(* CODESYS project process.library
   DefaultNamespace: KOSTAL.TC3.Core.process
   Description: Core Functionalities
   Author: Frank Dümpelmann
   DocFormat: reStructuredText
   Title: KOSTAL.TC3.Core.process
   Version: 2019.5.0.0
   Company: KOSTAL GmbH & Co.KG
   Placeholder: KOSTAL.TC3.Core.process

Project tree, tasks and I/O mapping:
  libraries: KOSTAL.TC3.Components.ListOf.Objects, 2019.1.0.0 (KOSTAL GmbH & Co.KG); KOSTAL.TC3.Components.Stringhandler, 2019.3.4.0 (KOSTAL GmbH & Co.KG); KOSTAL.TC3.Core.functionResponse, 2019.1.0.0 (KOSTAL GmbH & Co.KG); KOSTAL.TC3.Core.Settings, 2019.0.1.0 (KOSTAL GmbH & Co.KG); KOSTAL.TC3.Core.System, 2019.0.0.0 (KOSTAL GmbH & Co.KG)
  _Global/
    E_/
      data type E_PROCESS_CONDITION_DEFAULT_PRIORITYLEVEL
  Condition/
    DUT/
      ListOf/
        function block FB_ListOf_processCondition [ST]: _deletePayLoad, _Get_P, _New, Add_DUT, CopyFrom, CopyTo, Delete_DUT, Get_I, Get_IOwner
        interface I_ListOf_processCondition: CopyTo, Get_I
        interface I_ListOf_processCondition_CopyFrom: CopyFrom
        interface I_ListOf_processCondition_Owner: Add_DUT, CopyFrom, CopyTo, Delete_DUT, Get_I, Get_IOwner
      function block FB_processCondition [ST]: clear, CopyFrom, CopyTo, FB_init, getPriority, iMessage, isActive, isError, isInfo, isMasterMessage, isMessage, isText, message, PriorityLevel_Error, PriorityLevel_Info, PriorityLevel_MasterMessage, PriorityLevel_Message, PriorityLevel_Text, setMessage
      interface I_processCondition: getPriority, iMessage, isActive, isError, isInfo, isMasterMessage, isMessage, isText, PriorityLevel_Error, PriorityLevel_Info, PriorityLevel_MasterMessage, PriorityLevel_Message, PriorityLevel_Text
      interface I_processCondition_CopyFrom: CopyFrom
      interface I_processCondition_Owner: clear, CopyFrom, CopyTo, getPriority, iMessage, isActive, isError, isInfo, isMasterMessage, isMessage, isText, message, PriorityLevel_Error, PriorityLevel_Info, PriorityLevel_MasterMessage, PriorityLevel_Message, PriorityLevel_Text, setMessage
  Message/
    DUT/
      messageText/
        ListOf/
          function block FB_ListOf_messageText [ST]: _deletePayLoad, _Get_P, _New, Add_DUT, CopyFrom, CopyTo, Delete_DUT, Get_I, Get_IOwner
          interface I_ListOf_messageText: CopyTo, Get_I
          interface I_ListOf_messageText_CopyFrom: CopyFrom
          interface I_ListOf_messageText_Owner: Add_DUT, CopyFrom, CopyTo, Delete_DUT, Get_I, Get_IOwner
        function block FB_messageText [ST]: clear, CopyFrom, CopyTo, line_01, toString
        interface I_messageText: CopyTo, line_01, toString
        interface I_messageText_CopyFrom: CopyFrom
        interface I_messageText_Owner: clear, CopyFrom, CopyTo, line_01, toString
      messageText_2_lines/
        ListOf/
          function block FB_ListOf_messageText_2_lines [ST]: _deletePayLoad, _Get_P, _New, Add_DUT, CopyFrom, CopyTo, Delete_DUT, Get_I, Get_IOwner
          interface I_ListOf_messageText_2_lines: CopyTo, Get_I
          interface I_ListOf_messageText_2_lines_CopyFrom: CopyFrom
          interface I_ListOf_messageText_2_lines_Owner: Add_DUT, CopyFrom, CopyTo, Delete_DUT, Get_I, Get_IOwner
        function block FB_messageText_2_lines [ST]: clear, CopyFrom, line_02, toString
        interface I_messageText_2_lines: line_02
        interface I_messageText_2_lines_Owner: line_02
      messageText_3_lines/
        ListOf/
          function block FB_ListOf_messageText_3_lines [ST]: _deletePayLoad, _Get_P, _New, Add_DUT, CopyFrom, CopyTo, Delete_DUT, Get_I, Get_IOwner
          interface I_ListOf_messageText_3_lines: CopyTo, Get_I
          interface I_ListOf_messageText_3_lines_CopyFrom: CopyFrom
          interface I_ListOf_messageText_3_lines_Owner: Add_DUT, CopyFrom, CopyTo, Delete_DUT, Get_I, Get_IOwner
        function block FB_messageText_3_lines [ST]: clear, CopyFrom, line_03, toString
        interface I_messageText_3_lines: line_03
        interface I_messageText_3_lines_Owner: line_03
  Mode/
    DUT/
      ListOf/
        function block FB_ListOf_processMode [ST]: _deletePayLoad, _Get_P, _New, Add_DUT, CopyFrom, CopyTo, Delete_DUT, Get_I, Get_IOwner
        interface I_ListOf_processMode: CopyTo, Get_I
        interface I_ListOf_processMode_CopyFrom: CopyFrom
        interface I_ListOf_processMode_Owner: Add_DUT, CopyFrom, CopyTo, Delete_DUT, Get_I, Get_IOwner
      function block FB_processMode [ST]: automatic, clear, CopyFrom, CopyTo, manual
      interface I_processMode: automatic, CopyTo, manual
      interface I_processMode_CopyFrom: CopyFrom
      interface I_processMode_Owner: automatic, clear, CopyFrom, CopyTo, manual
  Project Information/
    function F_GetCompany [ST]
    function F_GetTitle [ST]
    function F_GetVersion [ST]
  State/
    DUT/
      ListOf/
        function block FB_ListOf_processState [ST]: _deletePayLoad, _Get_P, _New, Add_DUT, CopyFrom, CopyTo, Delete_DUT, Get_I, Get_IOwner
        interface I_ListOf_processState: CopyTo, Get_I
        interface I_ListOf_processState_CopyFrom: CopyFrom
        interface I_ListOf_processState_Owner: Add_DUT, CopyFrom, CopyTo, Delete_DUT, Get_I, Get_IOwner
      function block FB_processState [ST]: _clear_state, busy, calibrate, clear, CopyFrom, CopyTo, finish, off, on, ready, setUnique_busy, setUnique_calibrate, setUnique_finish, setUnique_off, setUnique_on, setUnique_ready
      interface I_processState: busy, calibrate, CopyTo, finish, off, on, ready
      interface I_processState_CopyFrom: CopyFrom
      interface I_processState_Owner: busy, calibrate, clear, CopyFrom, CopyTo, finish, off, on, ready, setUnique_busy, setUnique_calibrate, setUnique_finish, setUnique_off, setUnique_on, setUnique_ready
  Step/
    DUT/
      processStep/
        ListOf/
          function block FB_ListOf_processStep [ST]: _deletePayLoad, _Get_P, _New, Add_DUT, CopyFrom, CopyTo, Delete_DUT, Get_I, Get_IOwner
          interface I_ListOf_processStep: CopyTo, Get_I
          interface I_ListOf_processStep_CopyFrom: CopyFrom
          interface I_ListOf_processStep_Owner: Add_DUT, CopyFrom, CopyTo, Delete_DUT, Get_I, Get_IOwner
        function block FB_processStep [ST]: actual, clear, CopyFrom, CopyTo, DEC, Header, INC, init, request, set, toggle
        interface I_processStep: actual, CopyTo, request, toggle
        interface I_processStep_CopyFrom: CopyFrom
        interface I_processStep_Owner: actual, clear, CopyFrom, CopyTo, DEC, Header, INC, init, request, set, toggle
      processStep_Flow/
        ListOf/
          function block FB_ListOf_processStep_Flow [ST]: _deletePayLoad, _Get_P, _New, Add_DUT, CopyFrom, CopyTo, Delete_DUT, Get_I, Get_IOwner
          interface I_ListOf_processStep_Flow: CopyTo, Get_I
          interface I_ListOf_processStep_Flow_CopyFrom: CopyFrom
          interface I_ListOf_processStep_Flow_Owner: Add_DUT, CopyFrom, CopyTo, Delete_DUT, Get_I, Get_IOwner
        function block FB_processStep_Flow [ST]: clear, Header, init, isActive, isCalledExternally, NotFound
        interface I_processStep_Flow: isCalledExternally, NotFound
        interface I_processStep_Flow_Owner: clear, Header, init, isActive, isCalledExternally, NotFound
    GVL/
      global variables ProcessStep_GVL
    POE/
      ListOf/
        function block FB_ListOf_ProcessStep_Control [ST]: _deletePayLoad, _Get_P, _New, Add_DUT, CopyFrom, CopyTo, Delete_DUT, Get_I, Get_IOwner
        interface I_ListOf_ProcessStep_Control: CopyTo, Get_I
        interface I_ListOf_ProcessStep_Control_CopyFrom: CopyFrom
        interface I_ListOf_ProcessStep_Control_Owner: Add_DUT, CopyFrom, CopyTo, Delete_DUT, Get_I, Get_IOwner
      function block FB_ProcessStep_Control [ST]: _Forward, _modeAutomatik, _modeManual, BackwardDone, Condition, Control, CopyFrom, CopyTo, Done, ForwardDone, Header, iStep, JumpAddress, ManualBackward, ManualForward, ManualWithCondition, mode, Step
      interface I_ProcessStep_Control: BackwardDone, Condition, CopyTo, Done, ForwardDone, iStep, JumpAddress, ManualBackward, ManualForward, ManualWithCondition, mode
      interface I_ProcessStep_Control_CopyFrom: CopyFrom
      interface I_ProcessStep_Control_Owner: BackwardDone, Condition, Control, CopyFrom, CopyTo, Done, ForwardDone, Header, iStep, JumpAddress, ManualBackward, ManualForward, ManualWithCondition, mode, Step
  Version/
    global variables Global_Version
*)

// _Global/E_/E_PROCESS_CONDITION_DEFAULT_PRIORITYLEVEL
(*
Description
===========
| Levels of message priorities
| Intermediate values can be used to overrule other messages of the same level
| 1..999: INFORMATION - Display less important information (Color: grey)
| 1000..1999: TEXT_ONLY - To display information (Color: green)
| 2000..2999: MESSAGE - Order to the operator, e.g. 'Insert part' (Color: blue)
| 3000..3999: MASTERMESSAGE - Message to be displayed in upper HMI levels (Color: blue)
| 4000..4999: ERROR - Error message (Color: orange)

*)

{attribute 'qualified_only'}
TYPE E_PROCESS_CONDITION_DEFAULT_PRIORITYLEVEL :
(
	NONE 			:= 0,
	INFORMATION		:= 1,
	TEXT_ONLY		:= 1000,
	MESSAGE			:= 2000,
	MASTERMESSAGE	:= 3000,
	ERROR			:= 4000
);
END_TYPE

// Step/GVL/ProcessStep_GVL
{attribute 'qualified_only'}
VAR_GLOBAL CONSTANT
	PROCESS_STEP_INITIALIZE_STEP	: INT:= UINT_TO_INT(16#FFFF);
END_VAR

// Version/Global_Version
{attribute 'TcGenerated'}
{attribute 'no-analysis'}
{attribute 'linkalways'}
// This function has been automatically generated from the project information.
VAR_GLOBAL CONSTANT
	{attribute 'const_non_replaced'}
	stLibVersion_KOSTAL_TC3_Core_process : ST_LibVersion := (iMajor := 2019, iMinor := 5, iBuild := 0, iRevision := 0, nFlags := 1, sVersion := '2019.5.0.0');
END_VAR

// Condition/DUT/ListOf/FB_ListOf_processCondition
FUNCTION_BLOCK FB_ListOf_processCondition  EXTENDS KOSTAL_TC3_Components_ListOf_Objects.FB_Base IMPLEMENTS I_ListOf_processCondition, I_ListOf_processCondition_CopyFrom, I_ListOf_processCondition_Owner

VAR
	_Dummy	: FB_processCondition;
END_VAR

//Overwrites the method in the base class with the real contents of the ListOf class.
METHOD PROTECTED  _deletePayLoad
VAR_INPUT
	pPayload	:	PVOID; 
END_VAR

VAR
	_p	: POINTER TO FB_processCondition;
END_VAR

IF pPayload = 0  THEN	RETURN;	END_IF

_p:= pPayload;

__DELETE(_p);
END_METHOD

//Get read/write access to content
//Get_P returns a pointer to the Dummy instance
METHOD PROTECTED _Get_P : POINTER TO FB_processCondition

VAR_INPUT
	NumberOfObject	: UDINT;
	Response				: REFERENCE TO KOSTAL_TC3_Core_functionResponse.FB_functionResponse;
END_VAR

VAR
	_response: KOSTAL_TC3_Core_functionResponse.FB_functionResponse;
END_VAR

_response.clear();

IF (NumberOfObject = 0) 
OR (NumberOfObject > _ListOfObject.nObjects)
OR (_ListOfObject.pObjects = 0)
THEN

	_Dummy.Clear();

	_Get_P:= ADR(_Dummy);

	_response.status:= 'return Dummy because NumberOfPosition is out of range';

ELSE

	_response.success:= TRUE;
	
	_Get_P:= _ListOfObject.pObjects[NumberOfObject - 1];

END_IF

IF __ISVALIDREF(Response) THEN	Response.CopyFrom(_response);	END_IF
END_METHOD

//Overwrites the method in the base class with the real contents of the ListOf class.
METHOD PROTECTED  _New : PVOID

VAR
	_pNew: POINTER TO FB_processCondition;
END_VAR

_pNew:= __NEW(FB_processCondition);

_New:= _pNew;
END_METHOD

//Add a new instance of FB_Dut and copy content from [IN] to the new instance
METHOD PUBLIC Add_DUT : BOOL
VAR_INPUT
	IN				: I_processCondition;
	Response	: REFERENCE TO KOSTAL_TC3_Core_functionResponse.FB_functionResponse;
END_VAR

VAR
	pDUT: POINTER TO FB_processCondition;
	_response: KOSTAL_TC3_Core_functionResponse.FB_functionResponse;
END_VAR
_response.clear();

//create a new empty object 
IF NOT _AddObject() THEN
	_response.status:= ('_AddObject failed');
	IF __ISVALIDREF(Response) THEN	Response.CopyFrom(_response);	END_IF
	RETURN;	
END_IF

//Return, if no  [IN] object is available
IF IN = 0 THEN 
	_response.status:= ('IN Parameter not defined');
	IF __ISVALIDREF(Response) THEN	Response.CopyFrom(_response);	END_IF
	RETURN;	
END_IF

//otherwise fill [IN] object content to new virtual instance
pDUT:= _Get_P(_ListOfObject.nObjects, _response);

IF NOT _response.success THEN 
	IF __ISVALIDREF(Response) THEN	Response.CopyFrom(_response);	END_IF
	RETURN;	
END_IF

IF pDUT = 0 THEN 
	_response.status:= ('no Pointer get from list');
	IF __ISVALIDREF(Response) THEN	Response.CopyFrom(_response);	END_IF
	RETURN;	
END_IF

pDut^.CopyFrom(IN);

_response.success:= TRUE;
IF __ISVALIDREF(Response) THEN	Response.CopyFrom(_response);	END_IF

Add_DUT:= TRUE;
END_METHOD

METHOD PUBLIC CopyFrom
VAR_INPUT
	IN	: I_ListOf_processCondition;
END_VAR

VAR
	_udi: UDINT;
END_VAR

IF IN = 0 THEN RETURN;	END_IF

Clear();

FOR _udi:= 1 TO IN.NumberOfObjects DO
	Add_DUT(IN.Get_I(_udi, 0), 0);
END_FOR
END_METHOD

METHOD PUBLIC CopyTo
VAR_INPUT
	IN	: I_ListOf_processCondition_CopyFrom;
END_VAR

IF IN = 0 THEN RETURN;	END_IF

IN.CopyFrom(THIS^);
END_METHOD

METHOD PUBLIC Delete_DUT : BOOL
VAR_INPUT
	Number	: UDINT;	//Number of DUT in List
END_VAR

VAR
	_Set: FB_ListOf_processCondition;
	_udi: UDINT;
END_VAR

//Range control
IF Number = 0 							THEN RETURN;	END_IF
IF Number > NumberOfObjects	THEN RETURN;	END_IF

//Intermediate storage - prepare
_Set.Clear();

//catch all elements without the Number defiend
FOR _udi:= 1 TO NumberOfObjects DO
	IF _udi <> Number THEN
		_Set.Add_DUT(THIS^.Get_I(_udi, 0), 0);
	END_IF
END_FOR

//Delete own content
Clear();

//Add the remaining elements of the own class. 
FOR _udi:= 1 TO _Set.NumberOfObjects DO
		THIS^.Add_DUT(_Set.Get_I(_udi, 0), 0);
END_FOR

//Intermediate storage - clean Router storage
_Set.Clear();

Delete_DUT:= TRUE;
END_METHOD

//Get readonly access to content 
METHOD Get_I : I_processCondition

VAR_INPUT
	NumberOfObject	: UDINT;
	Response				: REFERENCE TO KOSTAL_TC3_Core_functionResponse.FB_functionResponse;
END_VAR

VAR
	_response: KOSTAL_TC3_Core_functionResponse.FB_functionResponse;
END_VAR

_response.clear();

Get_I:= _Get_P(NumberOfObject, _response)^;

IF __ISVALIDREF(Response) THEN	Response.CopyFrom(_response);	END_IF
END_METHOD

//Get readonly access to content 
METHOD Get_IOwner : I_processCondition_Owner

VAR_INPUT
	NumberOfObject	: UDINT;
	Response				: REFERENCE TO KOSTAL_TC3_Core_functionResponse.FB_functionResponse;
END_VAR

VAR
	_response: KOSTAL_TC3_Core_functionResponse.FB_functionResponse;
END_VAR

_response.clear();

Get_IOwner:= _Get_P(NumberOfObject, _response)^;

IF __ISVALIDREF(Response) THEN	Response.CopyFrom(_response);	END_IF
END_METHOD

END_FUNCTION_BLOCK

// Condition/DUT/ListOf/I_ListOf_processCondition
INTERFACE I_ListOf_processCondition EXTENDS KOSTAL_TC3_Components_ListOf_Objects.I_Base

METHOD PUBLIC CopyTo
VAR_INPUT
	IN	: I_ListOf_processCondition_CopyFrom;
END_VAR
END_METHOD

METHOD Get_I : I_processCondition

VAR_INPUT
	NumberOfObject	: UDINT;
	Response				: REFERENCE TO KOSTAL_TC3_Core_functionResponse.FB_functionResponse;
END_VAR
END_METHOD

END_INTERFACE

// Condition/DUT/ListOf/I_ListOf_processCondition_CopyFrom
INTERFACE I_ListOf_processCondition_CopyFrom EXTENDS KOSTAL_TC3_Core_System.I_Interface

METHOD PUBLIC CopyFrom
VAR_INPUT
	IN	: I_ListOf_processCondition;
END_VAR
END_METHOD

END_INTERFACE

// Condition/DUT/I_processCondition
INTERFACE I_processCondition EXTENDS KOSTAL_TC3_Core_System.I_Interface

METHOD PUBLIC getPriority : INT
VAR_INPUT
END_VAR
END_METHOD

(*
Description
===========
| Message to display in three lines
*)

PROPERTY PUBLIC iMessage : I_messageText_3_lines
GET
END_GET
END_PROPERTY

(*
Description
===========
| Returns TRUE if the user has a text, message or error to display
*)

METHOD PUBLIC isActive : BOOL
VAR_INPUT
END_VAR
END_METHOD

(*
Description
===========
| Returns TRUE if the user has an error to display
*)
METHOD PUBLIC isError : BOOL
VAR_INPUT
END_VAR
END_METHOD

(*
Description
===========
| Returns TRUE if the user has a message to display
*)
METHOD PUBLIC isInfo : BOOL
VAR_INPUT
END_VAR
END_METHOD

(*
Description
===========
| Returns TRUE if the user has a master message to display
*)
METHOD PUBLIC isMasterMessage : BOOL
VAR_INPUT
END_VAR
END_METHOD

(*
Description
===========
| Returns TRUE if the user has a message to display
*)
METHOD PUBLIC isMessage : BOOL
VAR_INPUT
END_VAR
END_METHOD

(*
Description
===========
| Returns TRUE if the user has a text to display
*)
METHOD PUBLIC isText : BOOL
END_METHOD

PROPERTY PUBLIC PriorityLevel_Error : INT
GET
END_GET
END_PROPERTY

PROPERTY PUBLIC PriorityLevel_Info : INT
GET
END_GET
END_PROPERTY

PROPERTY PUBLIC PriorityLevel_MasterMessage : INT
GET
END_GET
END_PROPERTY

PROPERTY PUBLIC PriorityLevel_Message : INT
GET
END_GET
END_PROPERTY

PROPERTY PUBLIC PriorityLevel_Text : INT
GET
END_GET
END_PROPERTY

END_INTERFACE

// Message/DUT/messageText_3_lines/I_messageText_3_lines
INTERFACE I_messageText_3_lines EXTENDS I_messageText_2_lines

PROPERTY PUBLIC line_03 : KOSTAL_TC3_Core_Settings.T_MaxString
GET
END_GET
END_PROPERTY

END_INTERFACE

// Message/DUT/messageText_2_lines/I_messageText_2_lines
INTERFACE I_messageText_2_lines EXTENDS I_messageText

PROPERTY PUBLIC line_02 : KOSTAL_TC3_Core_Settings.T_MaxString
GET
END_GET
END_PROPERTY

END_INTERFACE

// Message/DUT/messageText/I_messageText
INTERFACE I_messageText EXTENDS KOSTAL_TC3_Core_System.I_Interface

METHOD PUBLIC CopyTo
VAR_INPUT
	IN	:	I_messageText_CopyFrom;
END_VAR
END_METHOD

PROPERTY PUBLIC line_01 : KOSTAL_TC3_Core_Settings.T_MaxString
GET
END_GET
END_PROPERTY

METHOD PUBLIC toString : KOSTAL_TC3_Core_Settings.T_MaxString
END_METHOD

END_INTERFACE

// Message/DUT/messageText/I_messageText_CopyFrom
INTERFACE I_messageText_CopyFrom

METHOD PUBLIC CopyFrom
VAR_INPUT
	IN	: I_messageText;
END_VAR
END_METHOD

END_INTERFACE

// Condition/DUT/ListOf/I_ListOf_processCondition_Owner
INTERFACE I_ListOf_processCondition_Owner EXTENDS KOSTAL_TC3_Components_ListOf_Objects.I_Base_Owner

//Add a new instance of FB_Dut and copy content from [IN] to the new instance
METHOD PUBLIC Add_DUT : BOOL
VAR_INPUT
	IN				: I_processCondition;
	Response	: REFERENCE TO KOSTAL_TC3_Core_functionResponse.FB_functionResponse;
END_VAR
END_METHOD

METHOD PUBLIC CopyFrom
VAR_INPUT
	IN	: I_ListOf_processCondition;
END_VAR
END_METHOD

METHOD PUBLIC CopyTo
VAR_INPUT
	IN	: I_ListOf_processCondition_CopyFrom;
END_VAR
END_METHOD

METHOD PUBLIC Delete_DUT : BOOL
VAR_INPUT
	Number	: UDINT;	//Number of DUT in List
END_VAR
END_METHOD

METHOD Get_I : I_processCondition

VAR_INPUT
	NumberOfObject	: UDINT;
	Response				: REFERENCE TO KOSTAL_TC3_Core_functionResponse.FB_functionResponse;
END_VAR
END_METHOD

//Get readonly access to content 
METHOD Get_IOwner : I_processCondition_Owner

VAR_INPUT
	NumberOfObject	: UDINT;
	Response				: REFERENCE TO KOSTAL_TC3_Core_functionResponse.FB_functionResponse;
END_VAR
END_METHOD

END_INTERFACE

// Condition/DUT/I_processCondition_Owner
INTERFACE I_processCondition_Owner EXTENDS KOSTAL_TC3_Core_System.I_Interface

(*
Description
===========
| Clears existing message
*)

METHOD PUBLIC clear
END_METHOD

METHOD PUBLIC CopyFrom
VAR_INPUT
	IN	: I_processCondition;
END_VAR
END_METHOD

METHOD PUBLIC CopyTo
VAR_INPUT
	IN	:	I_processCondition_CopyFrom;
END_VAR
END_METHOD

METHOD PUBLIC getPriority : INT
VAR_INPUT
END_VAR
END_METHOD

(*
Description
===========
| Message to display in three lines
*)

PROPERTY PUBLIC iMessage : I_messageText_3_lines
GET
END_GET
END_PROPERTY

(*
Description
===========
| Returns TRUE if the user has a text, message or error to display
*)

METHOD PUBLIC isActive : BOOL
VAR_INPUT
END_VAR
END_METHOD

(*
Description
===========
| Returns TRUE if the user has an error to display
*)
METHOD PUBLIC isError : BOOL
VAR_INPUT
END_VAR
END_METHOD

(*
Description
===========
| Returns TRUE if the user has a message to display
*)
METHOD PUBLIC isInfo : BOOL
VAR_INPUT
END_VAR
END_METHOD

(*
Description
===========
| Returns TRUE if the user has a master message to display
*)
METHOD PUBLIC isMasterMessage : BOOL
VAR_INPUT
END_VAR
END_METHOD

(*
Description
===========
| Returns TRUE if the user has a message to display
*)
METHOD PUBLIC isMessage : BOOL
VAR_INPUT
END_VAR
END_METHOD

(*
Description
===========
| Returns TRUE if the user has a text to display
*)
METHOD PUBLIC isText : BOOL
END_METHOD

(*
Description
===========
| Message to display in three lines
*)

PROPERTY PUBLIC message : REFERENCE TO FB_messageText_3_lines
GET
END_GET
END_PROPERTY

PROPERTY PUBLIC PriorityLevel_Error : INT
GET
END_GET
END_PROPERTY

PROPERTY PUBLIC PriorityLevel_Info : INT
GET
END_GET
END_PROPERTY

PROPERTY PUBLIC PriorityLevel_MasterMessage : INT
GET
END_GET
END_PROPERTY

PROPERTY PUBLIC PriorityLevel_Message : INT
GET
END_GET
END_PROPERTY

PROPERTY PUBLIC PriorityLevel_Text : INT
GET
END_GET
END_PROPERTY

(*
Description
===========
| Sets message text and priority level for the user, in case the priority is higher than the existing message's priority 
| Existing messages with the same or lower priority are cleared
| Parameters:
| 	priority: INT - See E_PROCESS_CONDITION_DEFAULT_PRIORITYLEVEL for a detailed description
|	message: FB_messageText_3_lines - Content of the message
| Return value:
| 	FB_functionResponse: 
|		result: BOOL - Message ist set (no existing message with higher priority)
|		status: STRING(255) - Error description
*)

METHOD PUBLIC setMessage : FB_functionResponse

VAR_INPUT
	priority	: INT;
	message		: FB_messageText_3_lines;
END_VAR
END_METHOD

END_INTERFACE

// Condition/DUT/I_processCondition_CopyFrom
INTERFACE I_processCondition_CopyFrom EXTENDS KOSTAL_TC3_Core_System.I_Interface

METHOD PUBLIC CopyFrom
VAR_INPUT
	IN	: I_processCondition;
END_VAR
END_METHOD

END_INTERFACE

// Message/DUT/messageText_3_lines/FB_messageText_3_lines
(*

:Author: Frank Dümpelmann <f.duempelmann@kostal.com>
:Date: 2018-10-26

Function
========
| Data type containing three lines of text
| To be used in HMI communication

Methods and Properties
======================
| Clear(): Clears existing text
| line_01, line_02, line_03: Lines of text
*)

{attribute 'enable_dynamic_creation'}
FUNCTION_BLOCK PUBLIC FB_messageText_3_lines EXTENDS FB_messageText_2_lines IMPLEMENTS I_messageText_3_lines, I_messageText_3_lines_Owner

VAR
	_line_03	: KOSTAL_TC3_Core_Settings.T_MaxString;
END_VAR

(*
Description
===========
| Clears existing text
*)
METHOD PUBLIC clear
VAR_INPUT
END_VAR


SUPER^.clear();

_line_03:= '';
END_METHOD

METHOD PUBLIC CopyFrom
VAR_INPUT
	IN	: I_messageText;
END_VAR

VAR
	_obj		: I_messageText_3_lines;
	_bResult: BOOL;
END_VAR

IF IN = 0 THEN	RETURN;	END_IF

_bResult := __QUERYINTERFACE(IN, _obj);
 
IF NOT _bResult THEN RETURN;	END_IF
IF _obj = 0 THEN RETURN;	END_IF


SUPER^.CopyFrom(IN);
_line_03	:= _obj.line_03;
END_METHOD

PROPERTY PUBLIC line_03 : STRING(255)
GET

line_03:= _line_03;
END_GET
SET

_line_03:= line_03;
END_SET
END_PROPERTY

METHOD PUBLIC toString : STRING(255)

VAR
	_concat	: KOSTAL_TC3_Components_Stringhandler.FB_CONCAT;	//KOSTAL_TC3_Components_Stringhandler.FB_CONCAT
END_VAR

_concat.clear();
_concat.new(3);
_concat.addContent(1, SUPER^.toString());
_concat.addContent(2, ';');
_concat.addContent(3, _line_03);

toString:= _concat.getResult();
END_METHOD

END_FUNCTION_BLOCK

// Message/DUT/messageText_2_lines/FB_messageText_2_lines
(*

:Author: Frank Dümpelmann <f.duempelmann@kostal.com>
:Date: 2018-10-26

Function
========
| Data type containing two lines of text
| To be used in HMI communication

Methods and Properties
======================
| Clear(): Clears existing text
| line_01, line_02: Lines of text
*)

{attribute 'enable_dynamic_creation'}
FUNCTION_BLOCK PUBLIC FB_messageText_2_lines EXTENDS FB_messageText IMPLEMENTS I_messageText_2_lines, I_messageText_2_lines_Owner

VAR
	_line_02	: KOSTAL_TC3_Core_Settings.T_MaxString;
END_VAR

(*
Description
===========
| Clears existing text
*)
METHOD PUBLIC clear
VAR_INPUT
END_VAR


SUPER^.clear();

_line_02:= '';
END_METHOD

METHOD PUBLIC CopyFrom
VAR_INPUT
	IN	: I_messageText;
END_VAR

VAR
	_obj		: I_messageText_2_lines;
	_bResult: BOOL;
END_VAR

IF IN = 0 THEN	RETURN;	END_IF

_bResult := __QUERYINTERFACE(IN, _obj);
 
IF NOT _bResult THEN RETURN;	END_IF
IF _obj = 0 		THEN RETURN;	END_IF

SUPER^.CopyFrom(IN);
_line_02:= _obj.line_02;
END_METHOD

PROPERTY PUBLIC line_02 : KOSTAL_TC3_Core_Settings.T_MaxString
GET

line_02:= _line_02;
END_GET
SET

_line_02:= line_02;
END_SET
END_PROPERTY

METHOD PUBLIC toString : KOSTAL_TC3_Core_Settings.T_MaxString

VAR
	_concat	: KOSTAL_TC3_Components_Stringhandler.FB_CONCAT;	//KOSTAL_TC3_Components_Stringhandler.FB_CONCAT
END_VAR

_concat.clear();
_concat.new(3);
_concat.addContent(1, SUPER^.toString());
_concat.addContent(2, ';');
_concat.addContent(3, _line_02);

toString:= _concat.getResult();
END_METHOD

END_FUNCTION_BLOCK

// Message/DUT/messageText/FB_messageText
(*

:Author: Frank Dümpelmann <f.duempelmann@kostal.com>
:Date: 2018-10-26

Function
========
| Data type containing one line of text
| To be used in HMI communication

Methods and Properties
======================
| Clear(): Clears existing text
| line_01: Line of text
*)

{attribute 'enable_dynamic_creation'}
FUNCTION_BLOCK PUBLIC FB_messageText IMPLEMENTS I_messageText, I_messageText_CopyFrom, I_messageText_Owner

VAR
	_line_01	: KOSTAL_TC3_Core_Settings.T_MaxString;
END_VAR

(*
Description
===========
| Clears existing text
*)

METHOD PUBLIC clear
VAR_INPUT
END_VAR

_line_01:= '';
END_METHOD

METHOD PUBLIC CopyFrom
VAR_INPUT
	IN	: I_messageText;
END_VAR

IF IN = 0 THEN	RETURN;	END_IF

_line_01	:= IN.line_01;
END_METHOD

METHOD PUBLIC CopyTo
VAR_INPUT
	IN	:	I_messageText_CopyFrom;
END_VAR

IF IN = 0 THEN	RETURN;	END_IF

IN.CopyFrom(THIS^);
END_METHOD

PROPERTY PUBLIC line_01 : KOSTAL_TC3_Core_Settings.T_MaxString
GET

line_01:= _line_01;
END_GET
SET

_line_01:= line_01;
END_SET
END_PROPERTY

METHOD PUBLIC toString : KOSTAL_TC3_Core_Settings.T_MaxString

	
toString:= _line_01;
END_METHOD

END_FUNCTION_BLOCK

// Message/DUT/messageText/I_messageText_Owner
INTERFACE I_messageText_Owner EXTENDS KOSTAL_TC3_Core_System.I_Interface

(*
Description
===========
| Clears existing text
*)

METHOD PUBLIC clear
VAR_INPUT
END_VAR
END_METHOD

METHOD PUBLIC CopyFrom
VAR_INPUT
	IN	: I_messageText;
END_VAR
END_METHOD

METHOD PUBLIC CopyTo
VAR_INPUT
	IN	:	I_messageText_CopyFrom;
END_VAR
END_METHOD

PROPERTY PUBLIC line_01 : KOSTAL_TC3_Core_Settings.T_MaxString
GET
END_GET
SET
END_SET
END_PROPERTY

METHOD PUBLIC toString : KOSTAL_TC3_Core_Settings.T_MaxString
END_METHOD

END_INTERFACE

// Message/DUT/messageText_2_lines/I_messageText_2_lines_Owner
INTERFACE I_messageText_2_lines_Owner EXTENDS I_messageText_Owner

PROPERTY PUBLIC line_02 : KOSTAL_TC3_Core_Settings.T_MaxString
GET
END_GET
SET
END_SET
END_PROPERTY

END_INTERFACE

// Message/DUT/messageText_3_lines/I_messageText_3_lines_Owner
INTERFACE I_messageText_3_lines_Owner EXTENDS I_messageText_2_lines_Owner

PROPERTY PUBLIC line_03 : STRING(255)
GET
END_GET
SET
END_SET
END_PROPERTY

END_INTERFACE

// Condition/DUT/FB_processCondition
(*

:Author: Frank Dümpelmann <f.duempelmann@kostal.com>
:Date: 2018-10-26

Function
========
| Data structure representing the status of users/stations 
| Used for communication to superior instances, e.g. HMI

Usage notes
===============
| Call method setMessage from User/Station to set Message Text and priority level
| Call methods is... from the superior instance to get the user's status 
| Read message text from property message 

Methods and Properties
======================
| See bottom of this document for a detailed description of each method or property
*)

{attribute 'enable_dynamic_creation'}
FUNCTION_BLOCK PUBLIC FB_processCondition IMPLEMENTS I_processCondition, I_processCondition_CopyFrom, I_processCondition_Owner

VAR
	_priority	: INT;	//Priority of message
	
	_message	: FB_messageText_3_lines;
END_VAR

(*
Description
===========
| Clears existing message
*)

METHOD PUBLIC clear

_priority:= E_PROCESS_CONDITION_DEFAULT_PRIORITYLEVEL.NONE;

_message.clear();
END_METHOD

METHOD PUBLIC CopyFrom
VAR_INPUT
	IN	: I_processCondition;
END_VAR
IF IN = 0 THEN	RETURN;	END_IF

_message.CopyFrom(IN.iMessage);
END_METHOD

METHOD PUBLIC CopyTo
VAR_INPUT
	IN	:	I_processCondition_CopyFrom;
END_VAR

IF IN = 0 THEN	RETURN;	END_IF

IN.CopyFrom(THIS^);
END_METHOD

(*
Description
===========
| To be called automatically!
*)
METHOD FB_init : BOOL
VAR_INPUT
	bInitRetains : BOOL; // if TRUE, the retain variables are initialized (warm start / cold start)
	bInCopyCode : BOOL;  // if TRUE, the instance afterwards gets moved into the copy code (online change)
END_VAR
//_infoPriorityLevel			:= E_PROCESS_CONDITION_DEFAULT_PRIORITYLEVEL.INFORMATION; 
//_textPriorityLevel			:= E_PROCESS_CONDITION_DEFAULT_PRIORITYLEVEL.TEXT_ONLY;		//define the priority level from which priority a message is an user relative text 
//_messagePriorityLevel		:= E_PROCESS_CONDITION_DEFAULT_PRIORITYLEVEL.MESSAGE;		//define the priority level from which priority a message is an user relative message 
//_masterMessagePriorityLevel	:= E_PROCESS_CONDITION_DEFAULT_PRIORITYLEVEL.MASTERMESSAGE;	//define the priority level from which priority a message is an user relative error 
//_errorPriorityLevel			:= E_PROCESS_CONDITION_DEFAULT_PRIORITYLEVEL.ERROR;			//define the priority level from which priority a message is an user relative error
END_METHOD

METHOD PUBLIC getPriority : INT
VAR_INPUT
END_VAR

getPriority:= _priority;
END_METHOD

(*
Description
===========
| Message to display in three lines
*)

PROPERTY PUBLIC iMessage : I_messageText_3_lines
GET


iMessage := _message;
END_GET
END_PROPERTY

(*
Description
===========
| Returns TRUE if the user has a text, message or error to display
*)

METHOD PUBLIC isActive : BOOL
VAR_INPUT
END_VAR

isActive:= _priority <> E_PROCESS_CONDITION_DEFAULT_PRIORITYLEVEL.NONE;
END_METHOD

(*
Description
===========
| Returns TRUE if the user has an error to display
*)
METHOD PUBLIC isError : BOOL
VAR_INPUT
END_VAR

isError:= _priority >= E_PROCESS_CONDITION_DEFAULT_PRIORITYLEVEL.ERROR;
END_METHOD

(*
Description
===========
| Returns TRUE if the user has a message to display
*)
METHOD PUBLIC isInfo : BOOL
VAR_INPUT
END_VAR

isInfo:= (_priority >= E_PROCESS_CONDITION_DEFAULT_PRIORITYLEVEL.INFORMATION) AND (_priority < E_PROCESS_CONDITION_DEFAULT_PRIORITYLEVEL.TEXT_ONLY);
END_METHOD

(*
Description
===========
| Returns TRUE if the user has a master message to display
*)
METHOD PUBLIC isMasterMessage : BOOL
VAR_INPUT
END_VAR

isMasterMessage:= (_priority >= E_PROCESS_CONDITION_DEFAULT_PRIORITYLEVEL.MASTERMESSAGE) AND (_priority < E_PROCESS_CONDITION_DEFAULT_PRIORITYLEVEL.ERROR);
END_METHOD

(*
Description
===========
| Returns TRUE if the user has a message to display
*)
METHOD PUBLIC isMessage : BOOL
VAR_INPUT
END_VAR

isMessage:= (_priority >= E_PROCESS_CONDITION_DEFAULT_PRIORITYLEVEL.MESSAGE) AND (_priority < E_PROCESS_CONDITION_DEFAULT_PRIORITYLEVEL.MASTERMESSAGE);
END_METHOD

(*
Description
===========
| Returns TRUE if the user has a text to display
*)
METHOD PUBLIC isText : BOOL

isText:= (_priority >= E_PROCESS_CONDITION_DEFAULT_PRIORITYLEVEL.TEXT_ONLY) AND (_priority < E_PROCESS_CONDITION_DEFAULT_PRIORITYLEVEL.MESSAGE);
END_METHOD

(*
Description
===========
| Message to display in three lines
*)

PROPERTY PUBLIC message : REFERENCE TO FB_messageText_3_lines
GET


message REF= _message;
END_GET
END_PROPERTY

PROPERTY PUBLIC PriorityLevel_Error : INT
GET

PriorityLevel_Error := E_PROCESS_CONDITION_DEFAULT_PRIORITYLEVEL.ERROR;// _errorPriorityLevel;
END_GET
END_PROPERTY

PROPERTY PUBLIC PriorityLevel_Info : INT
GET

PriorityLevel_Info := E_PROCESS_CONDITION_DEFAULT_PRIORITYLEVEL.INFORMATION;
END_GET
END_PROPERTY

PROPERTY PUBLIC PriorityLevel_MasterMessage : INT
GET

PriorityLevel_MasterMessage := E_PROCESS_CONDITION_DEFAULT_PRIORITYLEVEL.MASTERMESSAGE;
END_GET
END_PROPERTY

PROPERTY PUBLIC PriorityLevel_Message : INT
GET

PriorityLevel_Message := E_PROCESS_CONDITION_DEFAULT_PRIORITYLEVEL.MESSAGE;
END_GET
END_PROPERTY

PROPERTY PUBLIC PriorityLevel_Text : INT
GET

PriorityLevel_Text := E_PROCESS_CONDITION_DEFAULT_PRIORITYLEVEL.TEXT_ONLY;
END_GET
END_PROPERTY

(*
Description
===========
| Sets message text and priority level for the user, in case the priority is higher than the existing message's priority 
| Existing messages with the same or lower priority are cleared
| Parameters:
| 	priority: INT - See E_PROCESS_CONDITION_DEFAULT_PRIORITYLEVEL for a detailed description
|	message: FB_messageText_3_lines - Content of the message
| Return value:
| 	FB_functionResponse: 
|		result: BOOL - Message ist set (no existing message with higher priority)
|		status: STRING(255) - Error description
*)

METHOD PUBLIC setMessage : FB_functionResponse

VAR_INPUT
	priority	: INT;
	message		: FB_messageText_3_lines;
END_VAR

IF priority > _priority THEN
	setMessage.clear();
	_priority	:= priority;
	_message	:= message;
	
	setMessage.Success	:= TRUE;

ELSE

	setMessage.Status	:= 'actual priority is higher';
	setMessage.Success	:= FALSE;

END_IF
END_METHOD

END_FUNCTION_BLOCK

// Message/DUT/messageText/ListOf/FB_ListOf_messageText
FUNCTION_BLOCK FB_ListOf_messageText  EXTENDS KOSTAL_TC3_Components_ListOf_Objects.FB_Base IMPLEMENTS I_ListOf_messageText, I_ListOf_messageText_CopyFrom, I_ListOf_messageText_Owner

VAR
	_Dummy	: FB_messageText;
END_VAR

//Overwrites the method in the base class with the real contents of the ListOf class.
METHOD PROTECTED  _deletePayLoad
VAR_INPUT
	pPayload	:	PVOID; 
END_VAR

VAR
	_p	: POINTER TO FB_messageText;
END_VAR

IF pPayload = 0  THEN	RETURN;	END_IF

_p:= pPayload;

__DELETE(_p);
END_METHOD

//Get read/write access to content
//Get_P returns a pointer to the Dummy instance
METHOD PROTECTED _Get_P : POINTER TO FB_messageText

VAR_INPUT
	NumberOfObject	: UDINT;
	Response				: REFERENCE TO KOSTAL_TC3_Core_functionResponse.FB_functionResponse;
END_VAR

VAR
	_response: KOSTAL_TC3_Core_functionResponse.FB_functionResponse;
END_VAR

_response.clear();

IF (NumberOfObject = 0) 
OR (NumberOfObject > _ListOfObject.nObjects)
OR (_ListOfObject.pObjects = 0)
THEN

	_Dummy.Clear();

	_Get_P:= ADR(_Dummy);

	_response.status:= 'return Dummy because NumberOfPosition is out of range';

ELSE

	_response.success:= TRUE;
	
	_Get_P:= _ListOfObject.pObjects[NumberOfObject - 1];

END_IF

IF __ISVALIDREF(Response) THEN	Response.CopyFrom(_response);	END_IF
END_METHOD

//Overwrites the method in the base class with the real contents of the ListOf class.
METHOD PROTECTED  _New : PVOID

VAR
	_pNew: POINTER TO FB_messageText;
END_VAR

_pNew:= __NEW(FB_messageText);

_New:= _pNew;
END_METHOD

//Add a new instance of FB_Dut and copy content from [IN] to the new instance
METHOD PUBLIC Add_DUT : BOOL
VAR_INPUT
	IN				: I_messageText;
	Response	: REFERENCE TO KOSTAL_TC3_Core_functionResponse.FB_functionResponse;
END_VAR

VAR
	pDUT: POINTER TO FB_messageText;
	_response: KOSTAL_TC3_Core_functionResponse.FB_functionResponse;
END_VAR
_response.clear();

//create a new empty object 
IF NOT _AddObject() THEN
	_response.status:= ('_AddObject failed');
	IF __ISVALIDREF(Response) THEN	Response.CopyFrom(_response);	END_IF
	RETURN;	
END_IF

//Return, if no  [IN] object is available
IF IN = 0 THEN 
	_response.status:= ('IN Parameter not defined');
	IF __ISVALIDREF(Response) THEN	Response.CopyFrom(_response);	END_IF
	RETURN;	
END_IF

//otherwise fill [IN] object content to new virtual instance
pDUT:= _Get_P(_ListOfObject.nObjects, _response);

IF NOT _response.success THEN 
	IF __ISVALIDREF(Response) THEN	Response.CopyFrom(_response);	END_IF
	RETURN;	
END_IF

IF pDUT = 0 THEN 
	_response.status:= ('no Pointer get from list');
	IF __ISVALIDREF(Response) THEN	Response.CopyFrom(_response);	END_IF
	RETURN;	
END_IF

pDut^.CopyFrom(IN);

_response.success:= TRUE;
IF __ISVALIDREF(Response) THEN	Response.CopyFrom(_response);	END_IF

Add_DUT:= TRUE;
END_METHOD

METHOD PUBLIC CopyFrom
VAR_INPUT
	IN	: I_ListOf_messageText;
END_VAR

VAR
	_udi: UDINT;
END_VAR

IF IN = 0 THEN RETURN;	END_IF

Clear();

FOR _udi:= 1 TO IN.NumberOfObjects DO
	Add_DUT(IN.Get_I(_udi, 0), 0);
END_FOR
END_METHOD

METHOD PUBLIC CopyTo
VAR_INPUT
	IN	: I_ListOf_messageText_CopyFrom;
END_VAR

IF IN = 0 THEN RETURN;	END_IF

IN.CopyFrom(THIS^);
END_METHOD

METHOD PUBLIC Delete_DUT : BOOL
VAR_INPUT
	Number	: UDINT;	//Number of DUT in List
END_VAR

VAR
	_Set: FB_ListOf_messageText;
	_udi: UDINT;
END_VAR

//Range control
IF Number = 0 							THEN RETURN;	END_IF
IF Number > NumberOfObjects	THEN RETURN;	END_IF

//Intermediate storage - prepare
_Set.Clear();

//catch all elements without the Number defiend
FOR _udi:= 1 TO NumberOfObjects DO
	IF _udi <> Number THEN
		_Set.Add_DUT(THIS^.Get_I(_udi, 0), 0);
	END_IF
END_FOR

//Delete own content
Clear();

//Add the remaining elements of the own class. 
FOR _udi:= 1 TO _Set.NumberOfObjects DO
		THIS^.Add_DUT(_Set.Get_I(_udi, 0), 0);
END_FOR

//Intermediate storage - clean Router storage
_Set.Clear();

Delete_DUT:= TRUE;
END_METHOD

//Get readonly access to content 
METHOD Get_I : I_messageText

VAR_INPUT
	NumberOfObject	: UDINT;
	Response				: REFERENCE TO KOSTAL_TC3_Core_functionResponse.FB_functionResponse;
END_VAR

VAR
	_response: KOSTAL_TC3_Core_functionResponse.FB_functionResponse;
END_VAR

_response.clear();

Get_I:= _Get_P(NumberOfObject, _response)^;

IF __ISVALIDREF(Response) THEN	Response.CopyFrom(_response);	END_IF
END_METHOD

//Get full access to content 
METHOD Get_IOwner : I_messageText_Owner

VAR_INPUT
	NumberOfObject	: UDINT;
	Response				: REFERENCE TO KOSTAL_TC3_Core_functionResponse.FB_functionResponse;
END_VAR

VAR
	_response: KOSTAL_TC3_Core_functionResponse.FB_functionResponse;
END_VAR

_response.clear();

Get_IOwner:= _Get_P(NumberOfObject, _response)^;

IF __ISVALIDREF(Response) THEN	Response.CopyFrom(_response);	END_IF
END_METHOD

END_FUNCTION_BLOCK

// Message/DUT/messageText/ListOf/I_ListOf_messageText
INTERFACE I_ListOf_messageText EXTENDS KOSTAL_TC3_Components_ListOf_Objects.I_Base

METHOD PUBLIC CopyTo
VAR_INPUT
	IN	: I_ListOf_messageText_CopyFrom;
END_VAR
END_METHOD

METHOD Get_I : I_messageText

VAR_INPUT
	NumberOfObject	: UDINT;
	Response				: REFERENCE TO KOSTAL_TC3_Core_functionResponse.FB_functionResponse;
END_VAR
END_METHOD

END_INTERFACE

// Message/DUT/messageText/ListOf/I_ListOf_messageText_CopyFrom
INTERFACE I_ListOf_messageText_CopyFrom EXTENDS KOSTAL_TC3_Core_System.I_Interface

METHOD PUBLIC CopyFrom
VAR_INPUT
	IN	: I_ListOf_messageText;
END_VAR
END_METHOD

END_INTERFACE

// Message/DUT/messageText/ListOf/I_ListOf_messageText_Owner
INTERFACE I_ListOf_messageText_Owner EXTENDS KOSTAL_TC3_Components_ListOf_Objects.I_Base_Owner

//Add a new instance of FB_Dut and copy content from [IN] to the new instance
METHOD PUBLIC Add_DUT : BOOL
VAR_INPUT
	IN				: I_messageText;
	Response	: REFERENCE TO KOSTAL_TC3_Core_functionResponse.FB_functionResponse;
END_VAR
END_METHOD

METHOD PUBLIC CopyFrom
VAR_INPUT
	IN	: I_ListOf_messageText;
END_VAR
END_METHOD

METHOD PUBLIC CopyTo
VAR_INPUT
	IN	: I_ListOf_messageText_CopyFrom;
END_VAR
END_METHOD

METHOD PUBLIC Delete_DUT : BOOL
VAR_INPUT
	Number	: UDINT;	//Number of DUT in List
END_VAR
END_METHOD

//Get readonly access to content 
METHOD Get_I : I_messageText

VAR_INPUT
	NumberOfObject	: UDINT;
	Response				: REFERENCE TO KOSTAL_TC3_Core_functionResponse.FB_functionResponse;
END_VAR
END_METHOD

//Get full access to content 
METHOD Get_IOwner : I_messageText_Owner

VAR_INPUT
	NumberOfObject	: UDINT;
	Response				: REFERENCE TO KOSTAL_TC3_Core_functionResponse.FB_functionResponse;
END_VAR
END_METHOD

END_INTERFACE

// Message/DUT/messageText_2_lines/ListOf/FB_ListOf_messageText_2_lines
FUNCTION_BLOCK FB_ListOf_messageText_2_lines  EXTENDS KOSTAL_TC3_Components_ListOf_Objects.FB_Base IMPLEMENTS I_ListOf_messageText_2_lines, I_ListOf_messageText_2_lines_CopyFrom, I_ListOf_messageText_2_lines_Owner

VAR
	_Dummy	: FB_messageText_2_lines;
END_VAR

//Overwrites the method in the base class with the real contents of the ListOf class.
METHOD PROTECTED  _deletePayLoad
VAR_INPUT
	pPayload	:	PVOID; 
END_VAR

VAR
	_p	: POINTER TO FB_messageText_2_lines;
END_VAR

IF pPayload = 0  THEN	RETURN;	END_IF

_p:= pPayload;

__DELETE(_p);
END_METHOD

//Get read/write access to content
//Get_P returns a pointer to the Dummy instance
METHOD PROTECTED _Get_P : POINTER TO FB_messageText_2_lines

VAR_INPUT
	NumberOfObject	: UDINT;
	Response				: REFERENCE TO KOSTAL_TC3_Core_functionResponse.FB_functionResponse;
END_VAR

VAR
	_response: KOSTAL_TC3_Core_functionResponse.FB_functionResponse;
END_VAR

_response.clear();

IF (NumberOfObject = 0) 
OR (NumberOfObject > _ListOfObject.nObjects)
OR (_ListOfObject.pObjects = 0)
THEN

	_Dummy.Clear();

	_Get_P:= ADR(_Dummy);

	_response.status:= 'return Dummy because NumberOfPosition is out of range';

ELSE

	_response.success:= TRUE;
	
	_Get_P:= _ListOfObject.pObjects[NumberOfObject - 1];

END_IF

IF __ISVALIDREF(Response) THEN	Response.CopyFrom(_response);	END_IF
END_METHOD

//Overwrites the method in the base class with the real contents of the ListOf class.
METHOD PROTECTED  _New : PVOID

VAR
	_pNew: POINTER TO FB_messageText_2_lines;
END_VAR

_pNew:= __NEW(FB_messageText_2_lines);

_New:= _pNew;
END_METHOD

//Add a new instance of FB_Dut and copy content from [IN] to the new instance
METHOD PUBLIC Add_DUT : BOOL
VAR_INPUT
	IN				: I_messageText_2_lines;
	Response	: REFERENCE TO KOSTAL_TC3_Core_functionResponse.FB_functionResponse;
END_VAR

VAR
	pDUT: POINTER TO FB_messageText_2_lines;
	_response: KOSTAL_TC3_Core_functionResponse.FB_functionResponse;
END_VAR
_response.clear();

//create a new empty object 
IF NOT _AddObject() THEN
	_response.status:= ('_AddObject failed');
	IF __ISVALIDREF(Response) THEN	Response.CopyFrom(_response);	END_IF
	RETURN;	
END_IF

//Return, if no  [IN] object is available
IF IN = 0 THEN 
	_response.status:= ('IN Parameter not defined');
	IF __ISVALIDREF(Response) THEN	Response.CopyFrom(_response);	END_IF
	RETURN;	
END_IF

//otherwise fill [IN] object content to new virtual instance
pDUT:= _Get_P(_ListOfObject.nObjects, _response);

IF NOT _response.success THEN 
	IF __ISVALIDREF(Response) THEN	Response.CopyFrom(_response);	END_IF
	RETURN;	
END_IF

IF pDUT = 0 THEN 
	_response.status:= ('no Pointer get from list');
	IF __ISVALIDREF(Response) THEN	Response.CopyFrom(_response);	END_IF
	RETURN;	
END_IF

pDut^.CopyFrom(IN);

_response.success:= TRUE;
IF __ISVALIDREF(Response) THEN	Response.CopyFrom(_response);	END_IF

Add_DUT:= TRUE;
END_METHOD

METHOD PUBLIC CopyFrom
VAR_INPUT
	IN	: I_ListOf_messageText_2_lines;
END_VAR

VAR
	_udi: UDINT;
END_VAR

IF IN = 0 THEN RETURN;	END_IF

Clear();

FOR _udi:= 1 TO IN.NumberOfObjects DO
	Add_DUT(IN.Get_I(_udi, 0), 0);
END_FOR
END_METHOD

METHOD PUBLIC CopyTo
VAR_INPUT
	IN	: I_ListOf_messageText_2_lines_CopyFrom;
END_VAR

IF IN = 0 THEN RETURN;	END_IF

IN.CopyFrom(THIS^);
END_METHOD

METHOD PUBLIC Delete_DUT : BOOL
VAR_INPUT
	Number	: UDINT;	//Number of DUT in List
END_VAR

VAR
	_Set: FB_ListOf_messageText_2_lines;
	_udi: UDINT;
END_VAR

//Range control
IF Number = 0 							THEN RETURN;	END_IF
IF Number > NumberOfObjects	THEN RETURN;	END_IF

//Intermediate storage - prepare
_Set.Clear();

//catch all elements without the Number defiend
FOR _udi:= 1 TO NumberOfObjects DO
	IF _udi <> Number THEN
		_Set.Add_DUT(THIS^.Get_I(_udi, 0), 0);
	END_IF
END_FOR

//Delete own content
Clear();

//Add the remaining elements of the own class. 
FOR _udi:= 1 TO _Set.NumberOfObjects DO
		THIS^.Add_DUT(_Set.Get_I(_udi, 0), 0);
END_FOR

//Intermediate storage - clean Router storage
_Set.Clear();

Delete_DUT:= TRUE;
END_METHOD

//Get readonly access to content 
METHOD Get_I : I_messageText_2_lines

VAR_INPUT
	NumberOfObject	: UDINT;
	Response				: REFERENCE TO KOSTAL_TC3_Core_functionResponse.FB_functionResponse;
END_VAR

VAR
	_response: KOSTAL_TC3_Core_functionResponse.FB_functionResponse;
END_VAR

_response.clear();

Get_I:= _Get_P(NumberOfObject, _response)^;

IF __ISVALIDREF(Response) THEN	Response.CopyFrom(_response);	END_IF
END_METHOD

//Get full access to content 
METHOD Get_IOwner : I_messageText_2_lines_Owner

VAR_INPUT
	NumberOfObject	: UDINT;
	Response				: REFERENCE TO KOSTAL_TC3_Core_functionResponse.FB_functionResponse;
END_VAR

VAR
	_response: KOSTAL_TC3_Core_functionResponse.FB_functionResponse;
END_VAR

_response.clear();

Get_IOwner:= _Get_P(NumberOfObject, _response)^;

IF __ISVALIDREF(Response) THEN	Response.CopyFrom(_response);	END_IF
END_METHOD

END_FUNCTION_BLOCK

// Message/DUT/messageText_2_lines/ListOf/I_ListOf_messageText_2_lines
INTERFACE I_ListOf_messageText_2_lines EXTENDS KOSTAL_TC3_Components_ListOf_Objects.I_Base

METHOD PUBLIC CopyTo
VAR_INPUT
	IN	: I_ListOf_messageText_2_lines_CopyFrom;
END_VAR
END_METHOD

METHOD Get_I : I_messageText_2_lines

VAR_INPUT
	NumberOfObject	: UDINT;
	Response				: REFERENCE TO KOSTAL_TC3_Core_functionResponse.FB_functionResponse;
END_VAR
END_METHOD

END_INTERFACE

// Message/DUT/messageText_2_lines/ListOf/I_ListOf_messageText_2_lines_CopyFrom
INTERFACE I_ListOf_messageText_2_lines_CopyFrom EXTENDS KOSTAL_TC3_Core_System.I_Interface

METHOD PUBLIC CopyFrom
VAR_INPUT
	IN	: I_ListOf_messageText_2_lines;
END_VAR
END_METHOD

END_INTERFACE

// Message/DUT/messageText_2_lines/ListOf/I_ListOf_messageText_2_lines_Owner
INTERFACE I_ListOf_messageText_2_lines_Owner EXTENDS KOSTAL_TC3_Components_ListOf_Objects.I_Base_Owner

//Add a new instance of FB_Dut and copy content from [IN] to the new instance
METHOD PUBLIC Add_DUT : BOOL
VAR_INPUT
	IN				: I_messageText_2_lines;
	Response	: REFERENCE TO KOSTAL_TC3_Core_functionResponse.FB_functionResponse;
END_VAR
END_METHOD

METHOD PUBLIC CopyFrom
VAR_INPUT
	IN	: I_ListOf_messageText_2_lines;
END_VAR
END_METHOD

METHOD PUBLIC CopyTo
VAR_INPUT
	IN	: I_ListOf_messageText_2_lines_CopyFrom;
END_VAR
END_METHOD

METHOD PUBLIC Delete_DUT : BOOL
VAR_INPUT
	Number	: UDINT;	//Number of DUT in List
END_VAR
END_METHOD

//Get readonly access to content 
METHOD Get_I : I_messageText_2_lines

VAR_INPUT
	NumberOfObject	: UDINT;
	Response				: REFERENCE TO KOSTAL_TC3_Core_functionResponse.FB_functionResponse;
END_VAR
END_METHOD

//Get full access to content 
METHOD Get_IOwner : I_messageText_2_lines_Owner

VAR_INPUT
	NumberOfObject	: UDINT;
	Response				: REFERENCE TO KOSTAL_TC3_Core_functionResponse.FB_functionResponse;
END_VAR
END_METHOD

END_INTERFACE

// Message/DUT/messageText_3_lines/ListOf/FB_ListOf_messageText_3_lines
FUNCTION_BLOCK FB_ListOf_messageText_3_lines  EXTENDS KOSTAL_TC3_Components_ListOf_Objects.FB_Base IMPLEMENTS I_ListOf_messageText_3_lines, I_ListOf_messageText_3_lines_CopyFrom, I_ListOf_messageText_3_lines_Owner

VAR
	_Dummy	: FB_messageText_3_lines;
END_VAR

//Overwrites the method in the base class with the real contents of the ListOf class.
METHOD PROTECTED  _deletePayLoad
VAR_INPUT
	pPayload	:	PVOID; 
END_VAR

VAR
	_p	: POINTER TO FB_messageText_3_lines;
END_VAR

IF pPayload = 0  THEN	RETURN;	END_IF

_p:= pPayload;

__DELETE(_p);
END_METHOD

//Get read/write access to content
//Get_P returns a pointer to the Dummy instance
METHOD PROTECTED _Get_P : POINTER TO FB_messageText_3_lines

VAR_INPUT
	NumberOfObject	: UDINT;
	Response				: REFERENCE TO KOSTAL_TC3_Core_functionResponse.FB_functionResponse;
END_VAR

VAR
	_response: KOSTAL_TC3_Core_functionResponse.FB_functionResponse;
END_VAR

_response.clear();

IF (NumberOfObject = 0) 
OR (NumberOfObject > _ListOfObject.nObjects)
OR (_ListOfObject.pObjects = 0)
THEN

	_Dummy.Clear();

	_Get_P:= ADR(_Dummy);

	_response.status:= 'return Dummy because NumberOfPosition is out of range';

ELSE

	_response.success:= TRUE;
	
	_Get_P:= _ListOfObject.pObjects[NumberOfObject - 1];

END_IF

IF __ISVALIDREF(Response) THEN	Response.CopyFrom(_response);	END_IF
END_METHOD

//Overwrites the method in the base class with the real contents of the ListOf class.
METHOD PROTECTED  _New : PVOID

VAR
	_pNew: POINTER TO FB_messageText_3_lines;
END_VAR

_pNew:= __NEW(FB_messageText_3_lines);

_New:= _pNew;
END_METHOD

//Add a new instance of FB_Dut and copy content from [IN] to the new instance
METHOD PUBLIC Add_DUT : BOOL
VAR_INPUT
	IN				: I_messageText_3_lines;
	Response	: REFERENCE TO KOSTAL_TC3_Core_functionResponse.FB_functionResponse;
END_VAR

VAR
	pDUT: POINTER TO FB_messageText_3_lines;
	_response: KOSTAL_TC3_Core_functionResponse.FB_functionResponse;
END_VAR
_response.clear();

//create a new empty object 
IF NOT _AddObject() THEN
	_response.status:= ('_AddObject failed');
	IF __ISVALIDREF(Response) THEN	Response.CopyFrom(_response);	END_IF
	RETURN;	
END_IF

//Return, if no  [IN] object is available
IF IN = 0 THEN 
	_response.status:= ('IN Parameter not defined');
	IF __ISVALIDREF(Response) THEN	Response.CopyFrom(_response);	END_IF
	RETURN;	
END_IF

//otherwise fill [IN] object content to new virtual instance
pDUT:= _Get_P(_ListOfObject.nObjects, _response);

IF NOT _response.success THEN 
	IF __ISVALIDREF(Response) THEN	Response.CopyFrom(_response);	END_IF
	RETURN;	
END_IF

IF pDUT = 0 THEN 
	_response.status:= ('no Pointer get from list');
	IF __ISVALIDREF(Response) THEN	Response.CopyFrom(_response);	END_IF
	RETURN;	
END_IF

pDut^.CopyFrom(IN);

_response.success:= TRUE;
IF __ISVALIDREF(Response) THEN	Response.CopyFrom(_response);	END_IF

Add_DUT:= TRUE;
END_METHOD

METHOD PUBLIC CopyFrom
VAR_INPUT
	IN	: I_ListOf_messageText_3_lines;
END_VAR

VAR
	_udi: UDINT;
END_VAR

IF IN = 0 THEN RETURN;	END_IF

Clear();

FOR _udi:= 1 TO IN.NumberOfObjects DO
	Add_DUT(IN.Get_I(_udi, 0), 0);
END_FOR
END_METHOD

METHOD PUBLIC CopyTo
VAR_INPUT
	IN	: I_ListOf_messageText_3_lines_CopyFrom;
END_VAR

IF IN = 0 THEN RETURN;	END_IF

IN.CopyFrom(THIS^);
END_METHOD

METHOD PUBLIC Delete_DUT : BOOL
VAR_INPUT
	Number	: UDINT;	//Number of DUT in List
END_VAR

VAR
	_Set: FB_ListOf_messageText_3_lines;
	_udi: UDINT;
END_VAR

//Range control
IF Number = 0 							THEN RETURN;	END_IF
IF Number > NumberOfObjects	THEN RETURN;	END_IF

//Intermediate storage - prepare
_Set.Clear();

//catch all elements without the Number defiend
FOR _udi:= 1 TO NumberOfObjects DO
	IF _udi <> Number THEN
		_Set.Add_DUT(THIS^.Get_I(_udi, 0), 0);
	END_IF
END_FOR

//Delete own content
Clear();

//Add the remaining elements of the own class. 
FOR _udi:= 1 TO _Set.NumberOfObjects DO
		THIS^.Add_DUT(_Set.Get_I(_udi, 0), 0);
END_FOR

//Intermediate storage - clean Router storage
_Set.Clear();

Delete_DUT:= TRUE;
END_METHOD

//Get readonly access to content 
METHOD Get_I : I_messageText_3_lines

VAR_INPUT
	NumberOfObject	: UDINT;
	Response				: REFERENCE TO KOSTAL_TC3_Core_functionResponse.FB_functionResponse;
END_VAR

VAR
	_response: KOSTAL_TC3_Core_functionResponse.FB_functionResponse;
END_VAR

_response.clear();

Get_I:= _Get_P(NumberOfObject, _response)^;

IF __ISVALIDREF(Response) THEN	Response.CopyFrom(_response);	END_IF
END_METHOD

//Get full access to content 
METHOD Get_IOwner : I_messageText_3_lines_Owner

VAR_INPUT
	NumberOfObject	: UDINT;
	Response				: REFERENCE TO KOSTAL_TC3_Core_functionResponse.FB_functionResponse;
END_VAR

VAR
	_response: KOSTAL_TC3_Core_functionResponse.FB_functionResponse;
END_VAR

_response.clear();

Get_IOwner:= _Get_P(NumberOfObject, _response)^;

IF __ISVALIDREF(Response) THEN	Response.CopyFrom(_response);	END_IF
END_METHOD

END_FUNCTION_BLOCK

// Message/DUT/messageText_3_lines/ListOf/I_ListOf_messageText_3_lines
INTERFACE I_ListOf_messageText_3_lines EXTENDS KOSTAL_TC3_Components_ListOf_Objects.I_Base

METHOD PUBLIC CopyTo
VAR_INPUT
	IN	: I_ListOf_messageText_3_lines_CopyFrom;
END_VAR
END_METHOD

METHOD Get_I : I_messageText_3_lines

VAR_INPUT
	NumberOfObject	: UDINT;
	Response				: REFERENCE TO KOSTAL_TC3_Core_functionResponse.FB_functionResponse;
END_VAR
END_METHOD

END_INTERFACE

// Message/DUT/messageText_3_lines/ListOf/I_ListOf_messageText_3_lines_CopyFrom
INTERFACE I_ListOf_messageText_3_lines_CopyFrom EXTENDS KOSTAL_TC3_Core_System.I_Interface

METHOD PUBLIC CopyFrom
VAR_INPUT
	IN	: I_ListOf_messageText_3_lines;
END_VAR
END_METHOD

END_INTERFACE

// Message/DUT/messageText_3_lines/ListOf/I_ListOf_messageText_3_lines_Owner
INTERFACE I_ListOf_messageText_3_lines_Owner EXTENDS KOSTAL_TC3_Components_ListOf_Objects.I_Base_Owner

//Add a new instance of FB_Dut and copy content from [IN] to the new instance
METHOD PUBLIC Add_DUT : BOOL
VAR_INPUT
	IN				: I_messageText_3_lines;
	Response	: REFERENCE TO KOSTAL_TC3_Core_functionResponse.FB_functionResponse;
END_VAR
END_METHOD

METHOD PUBLIC CopyFrom
VAR_INPUT
	IN	: I_ListOf_messageText_3_lines;
END_VAR
END_METHOD

METHOD PUBLIC CopyTo
VAR_INPUT
	IN	: I_ListOf_messageText_3_lines_CopyFrom;
END_VAR
END_METHOD

METHOD PUBLIC Delete_DUT : BOOL
VAR_INPUT
	Number	: UDINT;	//Number of DUT in List
END_VAR
END_METHOD

//Get readonly access to content 
METHOD Get_I : I_messageText_3_lines

VAR_INPUT
	NumberOfObject	: UDINT;
	Response				: REFERENCE TO KOSTAL_TC3_Core_functionResponse.FB_functionResponse;
END_VAR
END_METHOD

//Get full access to content 
METHOD Get_IOwner : I_messageText_3_lines_Owner

VAR_INPUT
	NumberOfObject	: UDINT;
	Response				: REFERENCE TO KOSTAL_TC3_Core_functionResponse.FB_functionResponse;
END_VAR
END_METHOD

END_INTERFACE

// Mode/DUT/ListOf/FB_ListOf_processMode
FUNCTION_BLOCK FB_ListOf_processMode  EXTENDS KOSTAL_TC3_Components_ListOf_Objects.FB_Base IMPLEMENTS I_ListOf_processMode, I_ListOf_processMode_CopyFrom, I_ListOf_processMode_Owner

VAR
	_Dummy	: FB_processMode;
END_VAR

//Overwrites the method in the base class with the real contents of the ListOf class.
METHOD PROTECTED  _deletePayLoad
VAR_INPUT
	pPayload	:	PVOID; 
END_VAR

VAR
	_p	: POINTER TO FB_processMode;
END_VAR

IF pPayload = 0  THEN	RETURN;	END_IF

_p:= pPayload;

__DELETE(_p);
END_METHOD

//Get read/write access to content
//Get_P returns a pointer to the Dummy instance
METHOD PROTECTED _Get_P : POINTER TO FB_processMode

VAR_INPUT
	NumberOfObject	: UDINT;
	Response				: REFERENCE TO KOSTAL_TC3_Core_functionResponse.FB_functionResponse;
END_VAR

VAR
	_response: KOSTAL_TC3_Core_functionResponse.FB_functionResponse;
END_VAR

_response.clear();

IF (NumberOfObject = 0) 
OR (NumberOfObject > _ListOfObject.nObjects)
OR (_ListOfObject.pObjects = 0)
THEN

	_Dummy.Clear();

	_Get_P:= ADR(_Dummy);

	_response.status:= 'return Dummy because NumberOfPosition is out of range';

ELSE

	_response.success:= TRUE;
	
	_Get_P:= _ListOfObject.pObjects[NumberOfObject - 1];

END_IF

IF __ISVALIDREF(Response) THEN	Response.CopyFrom(_response);	END_IF
END_METHOD

//Overwrites the method in the base class with the real contents of the ListOf class.
METHOD PROTECTED  _New : PVOID

VAR
	_pNew: POINTER TO FB_processMode;
END_VAR

_pNew:= __NEW(FB_processMode);

_New:= _pNew;
END_METHOD

//Add a new instance of FB_Dut and copy content from [IN] to the new instance
METHOD PUBLIC Add_DUT : BOOL
VAR_INPUT
	IN				: I_processMode;
	Response	: REFERENCE TO KOSTAL_TC3_Core_functionResponse.FB_functionResponse;
END_VAR

VAR
	pDUT: POINTER TO FB_processMode;
	_response: KOSTAL_TC3_Core_functionResponse.FB_functionResponse;
END_VAR
_response.clear();

//create a new empty object 
IF NOT _AddObject() THEN
	_response.status:= ('_AddObject failed');
	IF __ISVALIDREF(Response) THEN	Response.CopyFrom(_response);	END_IF
	RETURN;	
END_IF

//Return, if no  [IN] object is available
IF IN = 0 THEN 
	_response.status:= ('IN Parameter not defined');
	IF __ISVALIDREF(Response) THEN	Response.CopyFrom(_response);	END_IF
	RETURN;	
END_IF

//otherwise fill [IN] object content to new virtual instance
pDUT:= _Get_P(_ListOfObject.nObjects, _response);

IF NOT _response.success THEN 
	IF __ISVALIDREF(Response) THEN	Response.CopyFrom(_response);	END_IF
	RETURN;	
END_IF

IF pDUT = 0 THEN 
	_response.status:= ('no Pointer get from list');
	IF __ISVALIDREF(Response) THEN	Response.CopyFrom(_response);	END_IF
	RETURN;	
END_IF

pDut^.CopyFrom(IN);

_response.success:= TRUE;
IF __ISVALIDREF(Response) THEN	Response.CopyFrom(_response);	END_IF

Add_DUT:= TRUE;
END_METHOD

METHOD PUBLIC CopyFrom
VAR_INPUT
	IN	: I_ListOf_processMode;
END_VAR

VAR
	_udi: UDINT;
END_VAR

IF IN = 0 THEN RETURN;	END_IF

Clear();

FOR _udi:= 1 TO IN.NumberOfObjects DO
	Add_DUT(IN.Get_I(_udi, 0), 0);
END_FOR
END_METHOD

METHOD PUBLIC CopyTo
VAR_INPUT
	IN	: I_ListOf_processMode_CopyFrom;
END_VAR

IF IN = 0 THEN RETURN;	END_IF

IN.CopyFrom(THIS^);
END_METHOD

METHOD PUBLIC Delete_DUT : BOOL
VAR_INPUT
	Number	: UDINT;	//Number of DUT in List
END_VAR

VAR
	_Set: FB_ListOf_processMode;
	_udi: UDINT;
END_VAR

//Range control
IF Number = 0 							THEN RETURN;	END_IF
IF Number > NumberOfObjects	THEN RETURN;	END_IF

//Intermediate storage - prepare
_Set.Clear();

//catch all elements without the Number defiend
FOR _udi:= 1 TO NumberOfObjects DO
	IF _udi <> Number THEN
		_Set.Add_DUT(THIS^.Get_I(_udi, 0), 0);
	END_IF
END_FOR

//Delete own content
Clear();

//Add the remaining elements of the own class. 
FOR _udi:= 1 TO _Set.NumberOfObjects DO
		THIS^.Add_DUT(_Set.Get_I(_udi, 0), 0);
END_FOR

//Intermediate storage - clean Router storage
_Set.Clear();

Delete_DUT:= TRUE;
END_METHOD

//Get readonly access to content 
METHOD Get_I : I_processMode

VAR_INPUT
	NumberOfObject	: UDINT;
	Response				: REFERENCE TO KOSTAL_TC3_Core_functionResponse.FB_functionResponse;
END_VAR

VAR
	_response: KOSTAL_TC3_Core_functionResponse.FB_functionResponse;
END_VAR

_response.clear();

Get_I:= _Get_P(NumberOfObject, _response)^;

IF __ISVALIDREF(Response) THEN	Response.CopyFrom(_response);	END_IF
END_METHOD

//Get full access to content 
METHOD Get_IOwner : I_processMode_Owner

VAR_INPUT
	NumberOfObject	: UDINT;
	Response				: REFERENCE TO KOSTAL_TC3_Core_functionResponse.FB_functionResponse;
END_VAR

VAR
	_response: KOSTAL_TC3_Core_functionResponse.FB_functionResponse;
END_VAR

_response.clear();

Get_IOwner:= _Get_P(NumberOfObject, _response)^;

IF __ISVALIDREF(Response) THEN	Response.CopyFrom(_response);	END_IF
END_METHOD

END_FUNCTION_BLOCK

// Mode/DUT/ListOf/I_ListOf_processMode
INTERFACE I_ListOf_processMode EXTENDS KOSTAL_TC3_Components_ListOf_Objects.I_Base

METHOD PUBLIC CopyTo
VAR_INPUT
	IN	: I_ListOf_processMode_CopyFrom;
END_VAR
END_METHOD

METHOD Get_I : I_processMode

VAR_INPUT
	NumberOfObject	: UDINT;
	Response				: REFERENCE TO KOSTAL_TC3_Core_functionResponse.FB_functionResponse;
END_VAR
END_METHOD

END_INTERFACE

// Mode/DUT/ListOf/I_ListOf_processMode_CopyFrom
INTERFACE I_ListOf_processMode_CopyFrom EXTENDS KOSTAL_TC3_Core_System.I_Interface

METHOD PUBLIC CopyFrom
VAR_INPUT
	IN	: I_ListOf_processMode;
END_VAR
END_METHOD

END_INTERFACE

// Mode/DUT/I_processMode
INTERFACE I_processMode EXTENDS KOSTAL_TC3_Core_System.I_Interface

PROPERTY PUBLIC automatic : BOOL
GET
END_GET
END_PROPERTY

METHOD PUBLIC CopyTo
VAR_INPUT
	IN	:	I_processMode_CopyFrom;
END_VAR
END_METHOD

PROPERTY PUBLIC manual : BOOL
GET
END_GET
END_PROPERTY

END_INTERFACE

// Mode/DUT/I_processMode_CopyFrom
INTERFACE I_processMode_CopyFrom EXTENDS KOSTAL_TC3_Core_System.I_Interface

METHOD PUBLIC CopyFrom
VAR_INPUT
	IN	: I_processMode;
END_VAR
END_METHOD

END_INTERFACE

// Mode/DUT/ListOf/I_ListOf_processMode_Owner
INTERFACE I_ListOf_processMode_Owner EXTENDS KOSTAL_TC3_Components_ListOf_Objects.I_Base_Owner

//Add a new instance of FB_Dut and copy content from [IN] to the new instance
METHOD PUBLIC Add_DUT : BOOL
VAR_INPUT
	IN				: I_processMode;
	Response	: REFERENCE TO KOSTAL_TC3_Core_functionResponse.FB_functionResponse;
END_VAR
END_METHOD

METHOD PUBLIC CopyFrom
VAR_INPUT
	IN	: I_ListOf_processMode;
END_VAR
END_METHOD

METHOD PUBLIC CopyTo
VAR_INPUT
	IN	: I_ListOf_processMode_CopyFrom;
END_VAR
END_METHOD

METHOD PUBLIC Delete_DUT : BOOL
VAR_INPUT
	Number	: UDINT;	//Number of DUT in List
END_VAR
END_METHOD

//Get readonly access to content 
METHOD Get_I : I_processMode

VAR_INPUT
	NumberOfObject	: UDINT;
	Response				: REFERENCE TO KOSTAL_TC3_Core_functionResponse.FB_functionResponse;
END_VAR
END_METHOD

//Get full access to content 
METHOD Get_IOwner : I_processMode_Owner

VAR_INPUT
	NumberOfObject	: UDINT;
	Response				: REFERENCE TO KOSTAL_TC3_Core_functionResponse.FB_functionResponse;
END_VAR
END_METHOD

END_INTERFACE

// Mode/DUT/I_processMode_Owner
INTERFACE I_processMode_Owner EXTENDS KOSTAL_TC3_Core_System.I_Interface

PROPERTY PUBLIC automatic : BOOL
GET
END_GET
SET
END_SET
END_PROPERTY

METHOD PUBLIC clear
END_METHOD

METHOD PUBLIC CopyFrom
VAR_INPUT
	IN	: I_processMode;
END_VAR
END_METHOD

METHOD PUBLIC CopyTo
VAR_INPUT
	IN	:	I_processMode_CopyFrom;
END_VAR
END_METHOD

PROPERTY PUBLIC manual : BOOL
GET
END_GET
SET
END_SET
END_PROPERTY

END_INTERFACE

// Mode/DUT/FB_processMode
(*

:Author: Frank Dümpelmann <f.duempelmann@kostal.com>
:Date: 2018-10-26

Function
========
Data type representing the manual/automatic mode of an item
*)
{attribute 'enable_dynamic_creation'}
FUNCTION_BLOCK PUBLIC FB_processMode IMPLEMENTS I_processMode, I_processMode_CopyFrom, I_processMode_Owner

VAR
	_automatic	: BOOL;	//Release Automatic Functions
	_manual		: BOOL;	//Release Manual Functions	
END_VAR

PROPERTY PUBLIC automatic : BOOL
GET

automatic:= _automatic;
END_GET
SET

_automatic:= automatic;
END_SET
END_PROPERTY

METHOD PUBLIC clear

_automatic:= FALSE;
_manual		:= FALSE;
END_METHOD

METHOD PUBLIC CopyFrom
VAR_INPUT
	IN	: I_processMode;
END_VAR

IF IN = 0 THEN	RETURN;	END_IF

_automatic	:= IN.automatic;
_manual			:= IN.manual;
END_METHOD

METHOD PUBLIC CopyTo
VAR_INPUT
	IN	:	I_processMode_CopyFrom;
END_VAR

IF IN = 0 THEN	RETURN;	END_IF

IN.CopyFrom(THIS^);
END_METHOD

PROPERTY PUBLIC manual : BOOL
GET

manual:= _manual;
END_GET
SET

_manual:= manual;
END_SET
END_PROPERTY

END_FUNCTION_BLOCK

// Project Information/F_GetCompany
// This function has been automatically generated from the project information.
{attribute 'signature_flag' := '1073741824'}
{attribute 'TcGenerated'}
{attribute 'no-analysis'}
FUNCTION F_GetCompany : WSTRING
VAR_INPUT
	
END_VAR

F_GetCompany := "KOSTAL GmbH & Co.KG";

END_FUNCTION

// Project Information/F_GetTitle
// This function has been automatically generated from the project information.
{attribute 'signature_flag' := '1073741824'}
{attribute 'TcGenerated'}
{attribute 'no-analysis'}
FUNCTION F_GetTitle : WSTRING
VAR_INPUT
	
END_VAR

F_GetTitle := "KOSTAL.TC3.Core.process";

END_FUNCTION

// Project Information/F_GetVersion
// This function has been automatically generated from the project information.
{attribute 'signature_flag' := '1073741824'}
{attribute 'TcGenerated'}
{attribute 'no-analysis'}
FUNCTION F_GetVersion : ST_LibVersion
VAR_INPUT
	
END_VAR

F_GetVersion.iMajor := 2019;
F_GetVersion.iMinor := 5;
F_GetVersion.iBuild := 0;
F_GetVersion.iRevision := 0;
F_GetVersion.sVersion := '2019.5.0.0';
F_GetVersion.nFlags := 1;

END_FUNCTION

// State/DUT/ListOf/FB_ListOf_processState
FUNCTION_BLOCK FB_ListOf_processState  EXTENDS KOSTAL_TC3_Components_ListOf_Objects.FB_Base IMPLEMENTS I_ListOf_processState, I_ListOf_processState_CopyFrom, I_ListOf_processState_Owner

VAR
	_Dummy	: FB_processState;
END_VAR

//Overwrites the method in the base class with the real contents of the ListOf class.
METHOD PROTECTED  _deletePayLoad
VAR_INPUT
	pPayload	:	PVOID; 
END_VAR

VAR
	_p	: POINTER TO FB_processState;
END_VAR

IF pPayload = 0  THEN	RETURN;	END_IF

_p:= pPayload;

__DELETE(_p);
END_METHOD

//Get read/write access to content
//Get_P returns a pointer to the Dummy instance
METHOD PROTECTED _Get_P : POINTER TO FB_processState

VAR_INPUT
	NumberOfObject	: UDINT;
	Response				: REFERENCE TO KOSTAL_TC3_Core_functionResponse.FB_functionResponse;
END_VAR

VAR
	_response: KOSTAL_TC3_Core_functionResponse.FB_functionResponse;
END_VAR

_response.clear();

IF (NumberOfObject = 0) 
OR (NumberOfObject > _ListOfObject.nObjects)
OR (_ListOfObject.pObjects = 0)
THEN

	_Dummy.Clear();

	_Get_P:= ADR(_Dummy);

	_response.status:= 'return Dummy because NumberOfPosition is out of range';

ELSE

	_response.success:= TRUE;
	
	_Get_P:= _ListOfObject.pObjects[NumberOfObject - 1];

END_IF

IF __ISVALIDREF(Response) THEN	Response.CopyFrom(_response);	END_IF
END_METHOD

//Overwrites the method in the base class with the real contents of the ListOf class.
METHOD PROTECTED  _New : PVOID

VAR
	_pNew: POINTER TO FB_processState;
END_VAR

_pNew:= __NEW(FB_processState);

_New:= _pNew;
END_METHOD

//Add a new instance of FB_Dut and copy content from [IN] to the new instance
METHOD PUBLIC Add_DUT : BOOL
VAR_INPUT
	IN				: I_processState;
	Response	: REFERENCE TO KOSTAL_TC3_Core_functionResponse.FB_functionResponse;
END_VAR

VAR
	pDUT: POINTER TO FB_processState;
	_response: KOSTAL_TC3_Core_functionResponse.FB_functionResponse;
END_VAR
_response.clear();

//create a new empty object 
IF NOT _AddObject() THEN
	_response.status:= ('_AddObject failed');
	IF __ISVALIDREF(Response) THEN	Response.CopyFrom(_response);	END_IF
	RETURN;	
END_IF

//Return, if no  [IN] object is available
IF IN = 0 THEN 
	_response.status:= ('IN Parameter not defined');
	IF __ISVALIDREF(Response) THEN	Response.CopyFrom(_response);	END_IF
	RETURN;	
END_IF

//otherwise fill [IN] object content to new virtual instance
pDUT:= _Get_P(_ListOfObject.nObjects, _response);

IF NOT _response.success THEN 
	IF __ISVALIDREF(Response) THEN	Response.CopyFrom(_response);	END_IF
	RETURN;	
END_IF

IF pDUT = 0 THEN 
	_response.status:= ('no Pointer get from list');
	IF __ISVALIDREF(Response) THEN	Response.CopyFrom(_response);	END_IF
	RETURN;	
END_IF

pDut^.CopyFrom(IN);

_response.success:= TRUE;
IF __ISVALIDREF(Response) THEN	Response.CopyFrom(_response);	END_IF

Add_DUT:= TRUE;
END_METHOD

METHOD PUBLIC CopyFrom
VAR_INPUT
	IN	: I_ListOf_processState;
END_VAR

VAR
	_udi: UDINT;
END_VAR

IF IN = 0 THEN RETURN;	END_IF

Clear();

FOR _udi:= 1 TO IN.NumberOfObjects DO
	Add_DUT(IN.Get_I(_udi, 0), 0);
END_FOR
END_METHOD

METHOD PUBLIC CopyTo
VAR_INPUT
	IN	: I_ListOf_processState_CopyFrom;
END_VAR

IF IN = 0 THEN RETURN;	END_IF

IN.CopyFrom(THIS^);
END_METHOD

METHOD PUBLIC Delete_DUT : BOOL
VAR_INPUT
	Number	: UDINT;	//Number of DUT in List
END_VAR

VAR
	_Set: FB_ListOf_processState;
	_udi: UDINT;
END_VAR

//Range control
IF Number = 0 							THEN RETURN;	END_IF
IF Number > NumberOfObjects	THEN RETURN;	END_IF

//Intermediate storage - prepare
_Set.Clear();

//catch all elements without the Number defiend
FOR _udi:= 1 TO NumberOfObjects DO
	IF _udi <> Number THEN
		_Set.Add_DUT(THIS^.Get_I(_udi, 0), 0);
	END_IF
END_FOR

//Delete own content
Clear();

//Add the remaining elements of the own class. 
FOR _udi:= 1 TO _Set.NumberOfObjects DO
		THIS^.Add_DUT(_Set.Get_I(_udi, 0), 0);
END_FOR

//Intermediate storage - clean Router storage
_Set.Clear();

Delete_DUT:= TRUE;
END_METHOD

//Get readonly access to content 
METHOD Get_I : I_processState

VAR_INPUT
	NumberOfObject	: UDINT;
	Response				: REFERENCE TO KOSTAL_TC3_Core_functionResponse.FB_functionResponse;
END_VAR

VAR
	_response: KOSTAL_TC3_Core_functionResponse.FB_functionResponse;
END_VAR

_response.clear();

Get_I:= _Get_P(NumberOfObject, _response)^;

IF __ISVALIDREF(Response) THEN	Response.CopyFrom(_response);	END_IF
END_METHOD

//Get full access to content 
METHOD Get_IOwner : I_processState_Owner

VAR_INPUT
	NumberOfObject	: UDINT;
	Response				: REFERENCE TO KOSTAL_TC3_Core_functionResponse.FB_functionResponse;
END_VAR

VAR
	_response: KOSTAL_TC3_Core_functionResponse.FB_functionResponse;
END_VAR

_response.clear();

Get_IOwner:= _Get_P(NumberOfObject, _response)^;

IF __ISVALIDREF(Response) THEN	Response.CopyFrom(_response);	END_IF
END_METHOD

END_FUNCTION_BLOCK

// State/DUT/ListOf/I_ListOf_processState
INTERFACE I_ListOf_processState EXTENDS KOSTAL_TC3_Components_ListOf_Objects.I_Base

METHOD PUBLIC CopyTo
VAR_INPUT
	IN	: I_ListOf_processState_CopyFrom;
END_VAR
END_METHOD

METHOD Get_I : I_processState

VAR_INPUT
	NumberOfObject	: UDINT;
	Response				: REFERENCE TO KOSTAL_TC3_Core_functionResponse.FB_functionResponse;
END_VAR
END_METHOD

END_INTERFACE

// State/DUT/ListOf/I_ListOf_processState_CopyFrom
INTERFACE I_ListOf_processState_CopyFrom EXTENDS KOSTAL_TC3_Core_System.I_Interface

METHOD PUBLIC CopyFrom
VAR_INPUT
	IN	: I_ListOf_processState;
END_VAR
END_METHOD

END_INTERFACE

// State/DUT/I_processState
INTERFACE I_processState EXTENDS KOSTAL_TC3_Core_System.I_Interface

PROPERTY PUBLIC busy : BOOL
GET
END_GET
END_PROPERTY

PROPERTY PUBLIC calibrate : BOOL
GET
END_GET
END_PROPERTY

METHOD PUBLIC CopyTo
VAR_INPUT
	IN	:	I_processState_CopyFrom;
END_VAR
END_METHOD

PROPERTY PUBLIC finish : BOOL
GET
END_GET
END_PROPERTY

PROPERTY PUBLIC off : BOOL
GET
END_GET
END_PROPERTY

PROPERTY PUBLIC on : BOOL
GET
END_GET
END_PROPERTY

PROPERTY PUBLIC ready : BOOL
GET
END_GET
END_PROPERTY

END_INTERFACE

// State/DUT/I_processState_CopyFrom
INTERFACE I_processState_CopyFrom EXTENDS KOSTAL_TC3_Core_System.I_Interface

METHOD PUBLIC CopyFrom
VAR_INPUT
	IN	: I_processState;
END_VAR
END_METHOD

END_INTERFACE

// State/DUT/ListOf/I_ListOf_processState_Owner
INTERFACE I_ListOf_processState_Owner EXTENDS KOSTAL_TC3_Components_ListOf_Objects.I_Base_Owner

//Add a new instance of FB_Dut and copy content from [IN] to the new instance
METHOD PUBLIC Add_DUT : BOOL
VAR_INPUT
	IN				: I_processState;
	Response	: REFERENCE TO KOSTAL_TC3_Core_functionResponse.FB_functionResponse;
END_VAR
END_METHOD

METHOD PUBLIC CopyFrom
VAR_INPUT
	IN	: I_ListOf_processState;
END_VAR
END_METHOD

METHOD PUBLIC CopyTo
VAR_INPUT
	IN	: I_ListOf_processState_CopyFrom;
END_VAR
END_METHOD

METHOD PUBLIC Delete_DUT : BOOL
VAR_INPUT
	Number	: UDINT;	//Number of DUT in List
END_VAR
END_METHOD

//Get readonly access to content 
METHOD Get_I : I_processState

VAR_INPUT
	NumberOfObject	: UDINT;
	Response				: REFERENCE TO KOSTAL_TC3_Core_functionResponse.FB_functionResponse;
END_VAR
END_METHOD

//Get full access to content 
METHOD Get_IOwner : I_processState_Owner

VAR_INPUT
	NumberOfObject	: UDINT;
	Response				: REFERENCE TO KOSTAL_TC3_Core_functionResponse.FB_functionResponse;
END_VAR
END_METHOD

END_INTERFACE

// State/DUT/I_processState_Owner
INTERFACE I_processState_Owner EXTENDS KOSTAL_TC3_Core_System.I_Interface

PROPERTY PUBLIC busy : BOOL
GET
END_GET
SET
END_SET
END_PROPERTY

PROPERTY PUBLIC calibrate : BOOL
GET
END_GET
SET
END_SET
END_PROPERTY

METHOD PUBLIC clear
END_METHOD

METHOD PUBLIC CopyFrom
VAR_INPUT
	IN	: I_processState;
END_VAR
END_METHOD

METHOD PUBLIC CopyTo
VAR_INPUT
	IN	:	I_processState_CopyFrom;
END_VAR
END_METHOD

PROPERTY PUBLIC finish : BOOL
GET
END_GET
SET
END_SET
END_PROPERTY

PROPERTY PUBLIC off : BOOL
GET
END_GET
SET
END_SET
END_PROPERTY

PROPERTY PUBLIC on : BOOL
GET
END_GET
SET
END_SET
END_PROPERTY

PROPERTY PUBLIC ready : BOOL
GET
END_GET
SET
END_SET
END_PROPERTY

METHOD PUBLIC setUnique_busy
END_METHOD

METHOD PUBLIC setUnique_calibrate
END_METHOD

METHOD PUBLIC setUnique_finish
END_METHOD

METHOD PUBLIC setUnique_off
END_METHOD

METHOD PUBLIC setUnique_on
END_METHOD

METHOD PUBLIC setUnique_ready
END_METHOD

END_INTERFACE

// State/DUT/FB_processState
(*

:Author: Frank Dümpelmann <f.duempelmann@kostal.com>
:Date: 2018-10-26

Function
========
Data type representing the process state of an item

Methods and Properties
======================
| Properties represent the possible process states (off, on, calibrate, ready, busy, finish)
| Methods setUnique_... set the corresponding state and clear the others
| Alternatively, states can be set independent of the others using the properties 
| Methods starting with an underline(_) are internally used and can be ignored by the user
*)
{attribute 'enable_dynamic_creation'}
FUNCTION_BLOCK PUBLIC FB_processState IMPLEMENTS I_processState, I_processState_CopyFrom, I_processState_Owner

VAR
	_off 			: BOOL;	//BOOL
	_on 			: BOOL;	//BOOL
	_calibrate 		: BOOL;	//BOOL
	_ready 			: BOOL;	//BOOL
	_busy 			: BOOL;	//BOOL
	_finish 		: BOOL;	//BOOL
END_VAR

METHOD PROTECTED _clear_state

_busy		:= FALSE;
_calibrate	:= FALSE;
_finish		:= FALSE;
_off		:= FALSE;
_on			:= FALSE;
_ready		:= FALSE;
END_METHOD

PROPERTY PUBLIC busy : BOOL
GET

busy:= _busy;
END_GET
SET

_busy:= busy;
END_SET
END_PROPERTY

PROPERTY PUBLIC calibrate : BOOL
GET

calibrate:= _calibrate;
END_GET
SET

_calibrate:= calibrate;
END_SET
END_PROPERTY

METHOD PUBLIC clear

_clear_state();
END_METHOD

METHOD PUBLIC CopyFrom
VAR_INPUT
	IN	: I_processState;
END_VAR

IF IN = 0 THEN	RETURN;	END_IF

_busy				:= IN.busy;
_calibrate	:= IN.calibrate;
_finish			:= IN.finish;
_off				:= IN.off;
_on					:= IN.on;
_ready			:= IN.ready;
END_METHOD

METHOD PUBLIC CopyTo
VAR_INPUT
	IN	:	I_processState_CopyFrom;
END_VAR

IF IN = 0 THEN	RETURN;	END_IF

IN.CopyFrom(THIS^);
END_METHOD

PROPERTY PUBLIC finish : BOOL
GET

finish:= _finish;
END_GET
SET

_finish:= finish;
END_SET
END_PROPERTY

PROPERTY PUBLIC off : BOOL
GET

off:= _off;
END_GET
SET

_off:= off;
END_SET
END_PROPERTY

PROPERTY PUBLIC on : BOOL
GET

on:= _on;
END_GET
SET

_on:= on;
END_SET
END_PROPERTY

PROPERTY PUBLIC ready : BOOL
GET

ready:= _ready;
END_GET
SET

_ready:= ready;
END_SET
END_PROPERTY

METHOD PUBLIC setUnique_busy

_clear_state();

_busy:= TRUE;
END_METHOD

METHOD PUBLIC setUnique_calibrate

_clear_state();

_calibrate:= TRUE;
END_METHOD

METHOD PUBLIC setUnique_finish

_clear_state();

_finish:= TRUE;
END_METHOD

METHOD PUBLIC setUnique_off

_clear_state();

_off:= TRUE;
END_METHOD

METHOD PUBLIC setUnique_on

_clear_state();

_on:= TRUE;
END_METHOD

METHOD PUBLIC setUnique_ready

_clear_state();

_ready:= TRUE;
END_METHOD

END_FUNCTION_BLOCK

// Step/DUT/processStep/ListOf/FB_ListOf_processStep
FUNCTION_BLOCK FB_ListOf_processStep  EXTENDS KOSTAL_TC3_Components_ListOf_Objects.FB_Base IMPLEMENTS I_ListOf_processStep, I_ListOf_processStep_CopyFrom, I_ListOf_processStep_Owner

VAR
	_Dummy	: FB_processStep;
END_VAR

//Overwrites the method in the base class with the real contents of the ListOf class.
METHOD PROTECTED  _deletePayLoad
VAR_INPUT
	pPayload	:	PVOID; 
END_VAR

VAR
	_p	: POINTER TO FB_processStep;
END_VAR

IF pPayload = 0  THEN	RETURN;	END_IF

_p:= pPayload;

__DELETE(_p);
END_METHOD

//Get read/write access to content
//Get_P returns a pointer to the Dummy instance
METHOD PROTECTED _Get_P : POINTER TO FB_processStep

VAR_INPUT
	NumberOfObject	: UDINT;
	Response				: REFERENCE TO KOSTAL_TC3_Core_functionResponse.FB_functionResponse;
END_VAR

VAR
	_response: KOSTAL_TC3_Core_functionResponse.FB_functionResponse;
END_VAR

_response.clear();

IF (NumberOfObject = 0) 
OR (NumberOfObject > _ListOfObject.nObjects)
OR (_ListOfObject.pObjects = 0)
THEN

	_Dummy.Clear();

	_Get_P:= ADR(_Dummy);

	_response.status:= 'return Dummy because NumberOfPosition is out of range';

ELSE

	_response.success:= TRUE;
	
	_Get_P:= _ListOfObject.pObjects[NumberOfObject - 1];

END_IF

IF __ISVALIDREF(Response) THEN	Response.CopyFrom(_response);	END_IF
END_METHOD

//Overwrites the method in the base class with the real contents of the ListOf class.
METHOD PROTECTED  _New : PVOID

VAR
	_pNew: POINTER TO FB_processStep;
END_VAR

_pNew:= __NEW(FB_processStep);

_New:= _pNew;
END_METHOD

//Add a new instance of FB_Dut and copy content from [IN] to the new instance
METHOD PUBLIC Add_DUT : BOOL
VAR_INPUT
	IN				: I_processStep;
	Response	: REFERENCE TO KOSTAL_TC3_Core_functionResponse.FB_functionResponse;
END_VAR

VAR
	pDUT: POINTER TO FB_processStep;
	_response: KOSTAL_TC3_Core_functionResponse.FB_functionResponse;
END_VAR
_response.clear();

//create a new empty object 
IF NOT _AddObject() THEN
	_response.status:= ('_AddObject failed');
	IF __ISVALIDREF(Response) THEN	Response.CopyFrom(_response);	END_IF
	RETURN;	
END_IF

//Return, if no  [IN] object is available
IF IN = 0 THEN 
	_response.status:= ('IN Parameter not defined');
	IF __ISVALIDREF(Response) THEN	Response.CopyFrom(_response);	END_IF
	RETURN;	
END_IF

//otherwise fill [IN] object content to new virtual instance
pDUT:= _Get_P(_ListOfObject.nObjects, _response);

IF NOT _response.success THEN 
	IF __ISVALIDREF(Response) THEN	Response.CopyFrom(_response);	END_IF
	RETURN;	
END_IF

IF pDUT = 0 THEN 
	_response.status:= ('no Pointer get from list');
	IF __ISVALIDREF(Response) THEN	Response.CopyFrom(_response);	END_IF
	RETURN;	
END_IF

pDut^.CopyFrom(IN);

_response.success:= TRUE;
IF __ISVALIDREF(Response) THEN	Response.CopyFrom(_response);	END_IF

Add_DUT:= TRUE;
END_METHOD

METHOD PUBLIC CopyFrom
VAR_INPUT
	IN	: I_ListOf_processStep;
END_VAR

VAR
	_udi: UDINT;
END_VAR

IF IN = 0 THEN RETURN;	END_IF

Clear();

FOR _udi:= 1 TO IN.NumberOfObjects DO
	Add_DUT(IN.Get_I(_udi, 0), 0);
END_FOR
END_METHOD

METHOD PUBLIC CopyTo
VAR_INPUT
	IN	: I_ListOf_processStep_CopyFrom;
END_VAR

IF IN = 0 THEN RETURN;	END_IF

IN.CopyFrom(THIS^);
END_METHOD

METHOD PUBLIC Delete_DUT : BOOL
VAR_INPUT
	Number	: UDINT;	//Number of DUT in List
END_VAR

VAR
	_Set: FB_ListOf_processStep;
	_udi: UDINT;
END_VAR

//Range control
IF Number = 0 							THEN RETURN;	END_IF
IF Number > NumberOfObjects	THEN RETURN;	END_IF

//Intermediate storage - prepare
_Set.Clear();

//catch all elements without the Number defiend
FOR _udi:= 1 TO NumberOfObjects DO
	IF _udi <> Number THEN
		_Set.Add_DUT(THIS^.Get_I(_udi, 0), 0);
	END_IF
END_FOR

//Delete own content
Clear();

//Add the remaining elements of the own class. 
FOR _udi:= 1 TO _Set.NumberOfObjects DO
		THIS^.Add_DUT(_Set.Get_I(_udi, 0), 0);
END_FOR

//Intermediate storage - clean Router storage
_Set.Clear();

Delete_DUT:= TRUE;
END_METHOD

//Get readonly access to content 
METHOD Get_I : I_processStep

VAR_INPUT
	NumberOfObject	: UDINT;
	Response				: REFERENCE TO KOSTAL_TC3_Core_functionResponse.FB_functionResponse;
END_VAR

VAR
	_response: KOSTAL_TC3_Core_functionResponse.FB_functionResponse;
END_VAR

_response.clear();

Get_I:= _Get_P(NumberOfObject, _response)^;

IF __ISVALIDREF(Response) THEN	Response.CopyFrom(_response);	END_IF
END_METHOD

//Get full access to content 
METHOD Get_IOwner : I_processStep_Owner

VAR_INPUT
	NumberOfObject	: UDINT;
	Response				: REFERENCE TO KOSTAL_TC3_Core_functionResponse.FB_functionResponse;
END_VAR

VAR
	_response: KOSTAL_TC3_Core_functionResponse.FB_functionResponse;
END_VAR

_response.clear();

Get_IOwner:= _Get_P(NumberOfObject, _response)^;

IF __ISVALIDREF(Response) THEN	Response.CopyFrom(_response);	END_IF
END_METHOD

END_FUNCTION_BLOCK

// Step/DUT/processStep/ListOf/I_ListOf_processStep
INTERFACE I_ListOf_processStep EXTENDS KOSTAL_TC3_Components_ListOf_Objects.I_Base

METHOD PUBLIC CopyTo
VAR_INPUT
	IN	: I_ListOf_processStep_CopyFrom;
END_VAR
END_METHOD

METHOD Get_I : I_processStep

VAR_INPUT
	NumberOfObject	: UDINT;
	Response				: REFERENCE TO KOSTAL_TC3_Core_functionResponse.FB_functionResponse;
END_VAR
END_METHOD

END_INTERFACE

// Step/DUT/processStep/ListOf/I_ListOf_processStep_CopyFrom
INTERFACE I_ListOf_processStep_CopyFrom EXTENDS KOSTAL_TC3_Core_System.I_Interface

METHOD PUBLIC CopyFrom
VAR_INPUT
	IN	: I_ListOf_processStep;
END_VAR
END_METHOD

END_INTERFACE

// Step/DUT/processStep/I_processStep
INTERFACE I_processStep EXTENDS KOSTAL_TC3_Core_System.I_Interface

(*
Description
===========
| Actual step number
*)
PROPERTY PUBLIC actual : INT
GET
END_GET
END_PROPERTY

METHOD PUBLIC CopyTo
VAR_INPUT
	IN	:	I_processStep_CopyFrom;
END_VAR
END_METHOD

(*
Description
===========
| Requested step number (will be set with the next call of Header()
*)
PROPERTY PUBLIC request : INT
GET
END_GET
END_PROPERTY

(*
Description
===========
| Toggle signal for initialzation purposes
| Is set TRUE when Header() was called and the step number changed
| Is reset FALSE with the next call of Header() without changing step number
*)

PROPERTY PUBLIC toggle : BOOL
GET
END_GET
END_PROPERTY

END_INTERFACE

// Step/DUT/processStep/I_processStep_CopyFrom
INTERFACE I_processStep_CopyFrom EXTENDS KOSTAL_TC3_Core_System.I_Interface

METHOD PUBLIC CopyFrom
VAR_INPUT
	IN	: I_processStep;
END_VAR
END_METHOD

END_INTERFACE

// Step/DUT/processStep/ListOf/I_ListOf_processStep_Owner
INTERFACE I_ListOf_processStep_Owner EXTENDS KOSTAL_TC3_Components_ListOf_Objects.I_Base_Owner

//Add a new instance of FB_Dut and copy content from [IN] to the new instance
METHOD PUBLIC Add_DUT : BOOL
VAR_INPUT
	IN				: I_processStep;
	Response	: REFERENCE TO KOSTAL_TC3_Core_functionResponse.FB_functionResponse;
END_VAR
END_METHOD

METHOD PUBLIC CopyFrom
VAR_INPUT
	IN	: I_ListOf_processStep;
END_VAR
END_METHOD

METHOD PUBLIC CopyTo
VAR_INPUT
	IN	: I_ListOf_processStep_CopyFrom;
END_VAR
END_METHOD

METHOD PUBLIC Delete_DUT : BOOL
VAR_INPUT
	Number	: UDINT;	//Number of DUT in List
END_VAR
END_METHOD

//Get readonly access to content 
METHOD Get_I : I_processStep

VAR_INPUT
	NumberOfObject	: UDINT;
	Response				: REFERENCE TO KOSTAL_TC3_Core_functionResponse.FB_functionResponse;
END_VAR
END_METHOD

//Get full access to content 
METHOD Get_IOwner : I_processStep_Owner

VAR_INPUT
	NumberOfObject	: UDINT;
	Response				: REFERENCE TO KOSTAL_TC3_Core_functionResponse.FB_functionResponse;
END_VAR
END_METHOD

END_INTERFACE

// Step/DUT/processStep/I_processStep_Owner
INTERFACE I_processStep_Owner EXTENDS KOSTAL_TC3_Core_System.I_Interface

(*
Description
===========
| Actual step number
*)
PROPERTY PUBLIC actual : INT
GET
END_GET
SET
END_SET
END_PROPERTY

METHOD PUBLIC clear
END_METHOD

METHOD PUBLIC CopyFrom
VAR_INPUT
	IN	: I_processStep;
END_VAR
END_METHOD

METHOD PUBLIC CopyTo
VAR_INPUT
	IN	:	I_processStep_CopyFrom;
END_VAR
END_METHOD

(*
Description
===========
| Decrease step number by one (will be set with the next call of Header()
*)
METHOD DEC : KOSTAL_TC3_Core_functionResponse.FB_functionResponse
VAR_INPUT
END_VAR
END_METHOD

(*
Description
===========
| Apply changes in step sequence
| Call before or after the step sequence (see usage sample)
*)
METHOD PUBLIC Header
VAR_INPUT
END_VAR
END_METHOD

(*
Description
===========
| Increase step number by one (will be set with the next call of Header()
*)
METHOD INC : KOSTAL_TC3_Core_functionResponse.FB_functionResponse
VAR_INPUT
END_VAR
END_METHOD

(*
Description
===========
| Reset step sequence to 0
*)
METHOD PUBLIC init
END_METHOD

(*
Description
===========
| Requested step number (will be set with the next call of Header()
*)
PROPERTY PUBLIC request : INT
GET
END_GET
SET
END_SET
END_PROPERTY

(*
Description
===========
| Select step number (will be set with the next call of Header()
| Same function as property request
| Parameters:
| 	request: INT - step number to go to
*)
METHOD PUBLIC set

VAR_INPUT
	request	: INT;	//INT
END_VAR
END_METHOD

(*
Description
===========
| Toggle signal for initialzation purposes
| Is set TRUE when Header() was called and the step number changed
| Is reset FALSE with the next call of Header() without changing step number
*)

PROPERTY PUBLIC toggle : BOOL
GET
END_GET
SET
END_SET
END_PROPERTY

END_INTERFACE

// Step/DUT/processStep/FB_processStep
(*

:Author: Frank Dümpelmann <f.duempelmann@kostal.com>
:Date: 2018-10-26

Function
========
| Data structure representing a step sequence or state machine
| All changes are applied when the method Header() is called
| For the main step sequence of a station, use FB_ProcessStep_Control (implementig manual/automatic,...)

Methods and Properties
======================
| See bottom of this document for a detailed description of each method or property
| Methods starting with an underline(_) are internally used and can be ignored by the user

Usage sample:
=============

.. code:: 

	PROGRAM MAIN
	VAR
		_step : FB_processStep;
		_reset : BOOL := TRUE;
		_test1: BOOL;	
		_test2: INT;
		_test3: BOOL;
		_test4: BOOL;
	END_VAR
	
	IF _reset THEN
		_step.init();	//Init
		_reset := FALSE;
	END_IF
	
	_step.Header(); //Call before step sequence
	
	CASE _step.actual OF 
		0: 	IF (_test1) THEN
				_step.INC();	//Increase by one
			END_IF
		1: 	IF (_test2 > 1) THEN
				_step.request := 3;	//Set requested number directly
			ELSE
				_step.request := 4;	
			END_IF
		3: 	IF _test4 THEN
				_step.set(5);	//Set Method
			END_IF
			
		4: 	IF _test3 THEN
			_step.DEC();		//Decrease by one
			END_IF
		5: _reset := true;
	END_CASE
	
	IF _step.toggle THEN
	_toggleCounter := _toggleCounter+1;
	END_IF

*)

{attribute 'enable_dynamic_creation'}
FUNCTION_BLOCK FB_processStep IMPLEMENTS I_processStep, I_processStep_CopyFrom, I_processStep_Owner

VAR
	_actual		: INT;	//Actual Step Number
	_request	: INT;	//Requested Step Number
	_toggle		: BOOL;	//TRUE if actual Step Number is actualized with the requested
END_VAR

(*
Description
===========
| Actual step number
*)
PROPERTY PUBLIC actual : INT
GET

actual:= _actual;
END_GET
SET

_actual:= actual;
END_SET
END_PROPERTY

METHOD PUBLIC clear

_actual		:= 0;
_request	:= 0;
_toggle		:= FALSE;
END_METHOD

METHOD PUBLIC CopyFrom
VAR_INPUT
	IN	: I_processStep;
END_VAR

IF IN = 0 THEN	RETURN;	END_IF

_actual			:= IN.actual;
_request	:= IN.request;
_toggle		:= IN.toggle;
END_METHOD

METHOD PUBLIC CopyTo
VAR_INPUT
	IN	:	I_processStep_CopyFrom;
END_VAR

IF IN = 0 THEN	RETURN;	END_IF

IN.CopyFrom(THIS^);
END_METHOD

(*
Description
===========
| Decrease step number by one (will be set with the next call of Header()
*)
METHOD DEC : KOSTAL_TC3_Core_functionResponse.FB_functionResponse
VAR_INPUT
END_VAR


IF (_actual - 1) >  _actual THEN

	DEC.status	:= 'Overflow';
	DEC.success	:= FALSE;

ELSE

	_request:= _actual - 1;

	DEC.status	:= '';
	DEC.success	:= TRUE;
	
END_IF
END_METHOD

(*
Description
===========
| Apply changes in step sequence
| Call before or after the step sequence (see usage sample)
*)
METHOD PUBLIC Header
VAR_INPUT
END_VAR
_toggle:= _actual <> _request;
_actual := _request;
END_METHOD

(*
Description
===========
| Increase step number by one (will be set with the next call of Header()
*)
METHOD INC : KOSTAL_TC3_Core_functionResponse.FB_functionResponse
VAR_INPUT
END_VAR


IF (_actual + 1) <  _actual THEN

	INC.Status	:= 'Overflow';
	INC.Success	:= FALSE;

ELSE

	_request:= _actual + 1;

	INC.Status	:= '';
	INC.Success	:= TRUE;
	
END_IF
END_METHOD

(*
Description
===========
| Reset step sequence to 0
*)
METHOD PUBLIC init


_actual		:= UINT_TO_INT(16#FFFF);
_request	:= 0;
_toggle		:= TRUE;
END_METHOD

(*
Description
===========
| Requested step number (will be set with the next call of Header()
*)
PROPERTY PUBLIC request : INT
GET

request:= _request;
END_GET
SET

_request:= request;
END_SET
END_PROPERTY

(*
Description
===========
| Select step number (will be set with the next call of Header()
| Same function as property request
| Parameters:
| 	request: INT - step number to go to
*)
METHOD PUBLIC set

VAR_INPUT
	request	: INT;	//INT
END_VAR


_request:= request;
END_METHOD

(*
Description
===========
| Toggle signal for initialzation purposes
| Is set TRUE when Header() was called and the step number changed
| Is reset FALSE with the next call of Header() without changing step number
*)

PROPERTY PUBLIC toggle : BOOL
GET

toggle:= _toggle;
END_GET
SET

_toggle:= toggle;
END_SET
END_PROPERTY

END_FUNCTION_BLOCK

// Step/POE/FB_ProcessStep_Control
(*

:Author: Frank Dümpelmann <f.duempelmann@kostal.com>
:Date: 2018-10-26

Function
========
| Function block implementing the main step sequence of a station
| Variable step numbers, stepping forward and backward
| Feedback of successful step change
| Selection of manual or automatic stepping


Usage notes
===============
| Call method Header() before the step sequence
| Call method Control() at the end of each step to check the stepping condition 

Methods and Properties
======================
| See bottom of this document for a detailed description of each method or property
| Methods starting with an underline(_) are internally used and can be ignored by the user

Usage sample:
=============
| See framework or sample project MPL line

*)

{attribute 'enable_dynamic_creation'}
FUNCTION_BLOCK PUBLIC FB_ProcessStep_Control IMPLEMENTS I_ProcessStep_Control, I_ProcessStep_Control_CopyFrom, I_ProcessStep_Control_Owner

VAR
	_step	: FB_processStep;
	_mode	: FB_ProcessMode;	//ST_ProcessMode

	_condition						: BOOL;	//BOOL
	_manualWithCondition	: BOOL;	//BOOL
	_manualForward				: BOOL;	//BOOL
	_manualBackward				: BOOL;	//BOOL

	_jumpAddress					:	INT;	//INT

	_done					: BOOL;	//BOOL
	_backwardDone	: BOOL;	//BOOL
	_forwardDone	: BOOL;	//BOOL
	

END_VAR

METHOD PROTECTED _Forward : KOSTAL_TC3_Core_functionResponse.FB_functionResponse


	
IF _jumpAddress <> 0 THEN

	_step.set(_jumpAddress);

	_Forward.Status		:= '';
	_Forward.Success	:= TRUE;

	_jumpAddress:= 0;
	
ELSE

		_Forward:= _step.INC();

END_IF
END_METHOD

METHOD PROTECTED _modeAutomatik : KOSTAL_TC3_Core_functionResponse.FB_functionResponse

IF _condition THEN

	_condition:= FALSE;
	
	IF _jumpAddress <> 0 THEN

		_step.set(_jumpAddress);

		_done:= TRUE;	
		_jumpAddress:= 0;	
		
		_modeAutomatik.Status:= '';
		_modeAutomatik.Success:= TRUE;
		
	ELSE
		
		_modeAutomatik:= _step.INC();

		_done:= _modeAutomatik.Success;	
	
	END_IF
	
ELSE
	
	_modeAutomatik.Status:= 'Wait for condition';
	_modeAutomatik.Success:= TRUE;

END_IF
END_METHOD

METHOD PROTECTED _modeManual : KOSTAL_TC3_Core_functionResponse.FB_functionResponse


IF NOT _manualWithCondition OR _condition THEN

	_condition:= FALSE;
	
	IF _manualForward THEN

		_modeManual:= _Forward();
		
		IF _modeManual.Success THEN
			_manualForward	:= FALSE;
			_done						:= TRUE;	
			_forwardDone		:= TRUE;	
		END_IF

	ELSIF _manualBackward THEN

		
		_modeManual:=  _step.DEC();

		IF _modeManual.Success THEN	
			_manualBackward	:= FALSE;	
			_done						:= TRUE;	
			_backwardDone		:= TRUE;	
		END_IF

	ELSE

	_modeManual.Status:= 'Wait for manual request';
	_modeManual.Success:= TRUE;
		
	END_IF


ELSE
		
	_modeManual.Status:= 'Wait for condition';
	_modeManual.Success:= TRUE;

END_IF
END_METHOD

(*
Description
===========
| Step change backward was successful - Use e.g. to reset requests
| Attention: Variable is reset with next call of Header()
*)
PROPERTY PUBLIC BackwardDone : BOOL
GET

BackwardDone:= _backwardDone;

_backwardDone:= FALSE;
END_GET
END_PROPERTY

(*
Description
===========
| Condition to switch to the next step in automatic mode (also in manual mode if "ManualWithCondition" is TRUE) 
*)

PROPERTY PUBLIC Condition : BOOL
GET

Condition:= _condition;
END_GET
SET

_condition:= Condition;
END_SET
END_PROPERTY

(*
Description
===========
| Select next step number dependent of Condition and JumpAddress
*)

METHOD PUBLIC Control : FB_FunctionResponse

IF _mode.Automatic THEN
	
	Control := _modeAutomatik();

ELSIF _mode.Manual THEN

	Control := _modeManual();

ELSE

	Control.Status:= 'no mode detected';
	Control.Success:= TRUE;

END_IF
END_METHOD

METHOD PUBLIC CopyFrom
VAR_INPUT
	IN	: I_ProcessStep_Control;
END_VAR

IF IN = 0 THEN	RETURN;	END_IF

_backwardDone					:= IN.BackwardDone;
_condition						:= IN.Condition;
_done									:= IN.Done;
_forwardDone					:= IN.ForwardDone;
_jumpAddress					:= IN.JumpAddress;
_manualBackward				:= IN.ManualBackward;
_manualForward				:= IN.ManualForward;
_manualWithCondition	:= IN.ManualWithCondition;
_mode									:= IN.mode;

_step.CopyFrom(IN.iStep);
END_METHOD

METHOD PUBLIC CopyTo
VAR_INPUT
	IN	:	I_ProcessStep_Control_CopyFrom;
END_VAR

IF IN = 0 THEN	RETURN;	END_IF

IN.CopyFrom(THIS^);
END_METHOD

(*
Description
===========
| Step change was successful - Use e.g. to reset requests
| Attention: Variable is reset with next call of Header()
*)
PROPERTY PUBLIC Done : BOOL
GET

Done:= _done;

_done:= FALSE;
END_GET
END_PROPERTY

(*
Description
===========
| Step change forward was successful - Use e.g. to reset requests
| Attention: Variable is reset with next call of Header()
*)
PROPERTY PUBLIC ForwardDone : BOOL
GET

ForwardDone:= _forwardDone;

_forwardDone:= FALSE;
END_GET
END_PROPERTY

(*
Description
===========
| Apply changes in step sequence
| Call before the step sequence (see usage sample)
*)
METHOD PUBLIC Header

_step.Header();


_done			:= FALSE;
_backwardDone	:= FALSE;
_forwardDone	:= FALSE;
END_METHOD

(*
Description
===========
| FB_processStep containing the step data of the step control
| Full access to all parameters
| See documentation of FB_processStep for details

*)
PROPERTY PUBLIC iStep : I_processStep
GET

iStep:= _step;
END_GET
END_PROPERTY

(*
Description
===========
| Step number to go to next
| 0 = subsequent step
*)
PROPERTY PUBLIC JumpAddress : INT
GET


JumpAddress:= _jumpAddress;
END_GET
SET

_jumpAddress:= JumpAddress;
END_SET
END_PROPERTY

(*
Description
===========
| Go one step back in manual mode(pulse input - Backward button on HMI): 
*)
PROPERTY PUBLIC ManualBackward : BOOL
GET

ManualBackward:= _manualBackward;
END_GET
SET

_manualBackward:= ManualBackward;
END_SET
END_PROPERTY

(*
Description
===========
| Go to the next step (JumpAddress) in manual mode(pulse input - Forward button on HMI)
*)
PROPERTY PUBLIC ManualForward : BOOL
GET

ManualForward:= _manualForward;
END_GET
SET

_manualForward:= ManualForward;
END_SET
END_PROPERTY

(*
Description
===========
| If TRUE, property "Condition" is also active in manual mode
*)
PROPERTY PUBLIC ManualWithCondition : BOOL
GET

ManualWithCondition:= _manualWithCondition;
END_GET
SET

_manualWithCondition:= ManualWithCondition;
END_SET
END_PROPERTY

(*
Description
===========
| automatic: Control automatically jumps to the next step if Condition is TRUE
| manual: Input ManualForward must be pulsed TRUE to go to the next step
*)
PROPERTY PUBLIC mode : REFERENCE to FB_processMode
GET

mode REF= _mode;
END_GET
SET

_mode := mode;
END_SET
END_PROPERTY

(*
Description
===========
| FB_processStep containing the step data of the step control
| Full access to all parameters
| See documentation of FB_processStep for details

*)
PROPERTY PUBLIC Step : REFERENCE TO FB_processStep
GET

Step REF= _step;
END_GET
END_PROPERTY

END_FUNCTION_BLOCK

// Step/POE/I_ProcessStep_Control
(*

:Author: Martin Hundt <m.hundt@kostal.com>
:Date: 2019-04-18

Function
========
Interface to link current state/content from FB_ProcessStep_Control to other components which analyse the step sequence internally (e.g. FB_Cylinder_Controlled)
*)
INTERFACE I_ProcessStep_Control EXTENDS KOSTAL_TC3_Core_System.I_Interface

(*
Description
===========
| Step change backward was successful - Use e.g. to reset requests
| Attention: Variable is reset with next call of Header()
*)
PROPERTY PUBLIC BackwardDone : BOOL
GET
END_GET
END_PROPERTY

(*
Description
===========
| Condition to switch to the next step in automatic mode (also in manual mode if "ManualWithCondition" is TRUE) 
*)

PROPERTY PUBLIC Condition : BOOL
GET
END_GET
END_PROPERTY

METHOD PUBLIC CopyTo
VAR_INPUT
	IN	:	I_ProcessStep_Control_CopyFrom;
END_VAR
END_METHOD

(*
Description
===========
| Step change was successful - Use e.g. to reset requests
| Attention: Variable is reset with next call of Header()
*)
PROPERTY PUBLIC Done : BOOL
GET
END_GET
END_PROPERTY

(*
Description
===========
| Step change forward was successful - Use e.g. to reset requests
| Attention: Variable is reset with next call of Header()
*)
PROPERTY PUBLIC ForwardDone : BOOL
GET
END_GET
END_PROPERTY

(*
Description
===========
| FB_processStep containing the step data of the step control
| Full access to all parameters
| See documentation of FB_processStep for details

*)
PROPERTY PUBLIC iStep : I_processStep
GET
END_GET
END_PROPERTY

(*
Description
===========
| Step number to go to next
| 0 = subsequent step
*)
PROPERTY PUBLIC JumpAddress : INT
GET
END_GET
END_PROPERTY

(*
Description
===========
| Go one step back in manual mode(pulse input - Backward button on HMI): 
*)
PROPERTY PUBLIC ManualBackward : BOOL
GET
END_GET
END_PROPERTY

(*
Description
===========
| Go to the next step (JumpAddress) in manual mode(pulse input - Forward button on HMI)
*)
PROPERTY PUBLIC ManualForward : BOOL
GET
END_GET
END_PROPERTY

(*
Description
===========
| If TRUE, property "Condition" is also active in manual mode
*)
PROPERTY PUBLIC ManualWithCondition : BOOL
GET
END_GET
END_PROPERTY

(*
Description
===========
| automatic: Control automatically jumps to the next step if Condition is TRUE
| manual: Input ManualForward must be pulsed TRUE to go to the next step
*)
PROPERTY PUBLIC mode : REFERENCE to FB_processMode
GET
END_GET
END_PROPERTY

END_INTERFACE

// Step/POE/I_ProcessStep_Control_CopyFrom
INTERFACE I_ProcessStep_Control_CopyFrom EXTENDS KOSTAL_TC3_Core_System.I_Interface

METHOD PUBLIC CopyFrom
VAR_INPUT
	IN	: I_ProcessStep_Control;
END_VAR
END_METHOD

END_INTERFACE

// Step/POE/I_ProcessStep_Control_Owner
INTERFACE I_ProcessStep_Control_Owner EXTENDS KOSTAL_TC3_Core_System.I_Interface

(*
Description
===========
| Step change backward was successful - Use e.g. to reset requests
| Attention: Variable is reset with next call of Header()
*)
PROPERTY PUBLIC BackwardDone : BOOL
GET
END_GET
END_PROPERTY

(*
Description
===========
| Condition to switch to the next step in automatic mode (also in manual mode if "ManualWithCondition" is TRUE) 
*)

PROPERTY PUBLIC Condition : BOOL
GET
END_GET
SET
END_SET
END_PROPERTY

(*
Description
===========
| Select next step number dependent of Condition and JumpAddress
*)

METHOD PUBLIC Control : FB_FunctionResponse
END_METHOD

METHOD PUBLIC CopyFrom
VAR_INPUT
	IN	: I_ProcessStep_Control;
END_VAR
END_METHOD

METHOD PUBLIC CopyTo
VAR_INPUT
	IN	:	I_ProcessStep_Control_CopyFrom;
END_VAR
END_METHOD

(*
Description
===========
| Step change was successful - Use e.g. to reset requests
| Attention: Variable is reset with next call of Header()
*)
PROPERTY PUBLIC Done : BOOL
GET
END_GET
END_PROPERTY

(*
Description
===========
| Step change forward was successful - Use e.g. to reset requests
| Attention: Variable is reset with next call of Header()
*)
PROPERTY PUBLIC ForwardDone : BOOL
GET
END_GET
END_PROPERTY

(*
Description
===========
| Apply changes in step sequence
| Call before the step sequence (see usage sample)
*)
METHOD PUBLIC Header
END_METHOD

(*
Description
===========
| FB_processStep containing the step data of the step control
| Full access to all parameters
| See documentation of FB_processStep for details

*)
PROPERTY PUBLIC iStep : I_processStep
GET
END_GET
END_PROPERTY

(*
Description
===========
| Step number to go to next
| 0 = subsequent step
*)
PROPERTY PUBLIC JumpAddress : INT
GET
END_GET
SET
END_SET
END_PROPERTY

(*
Description
===========
| Go one step back in manual mode(pulse input - Backward button on HMI): 
*)
PROPERTY PUBLIC ManualBackward : BOOL
GET
END_GET
SET
END_SET
END_PROPERTY

(*
Description
===========
| Go to the next step (JumpAddress) in manual mode(pulse input - Forward button on HMI)
*)
PROPERTY PUBLIC ManualForward : BOOL
GET
END_GET
SET
END_SET
END_PROPERTY

(*
Description
===========
| If TRUE, property "Condition" is also active in manual mode
*)
PROPERTY PUBLIC ManualWithCondition : BOOL
GET
END_GET
SET
END_SET
END_PROPERTY

(*
Description
===========
| automatic: Control automatically jumps to the next step if Condition is TRUE
| manual: Input ManualForward must be pulsed TRUE to go to the next step
*)
PROPERTY PUBLIC mode : REFERENCE to FB_processMode
GET
END_GET
SET
END_SET
END_PROPERTY

(*
Description
===========
| FB_processStep containing the step data of the step control
| Full access to all parameters
| See documentation of FB_processStep for details

*)
PROPERTY PUBLIC Step : REFERENCE TO FB_processStep
GET
END_GET
END_PROPERTY

END_INTERFACE

// Step/DUT/processStep_Flow/ListOf/FB_ListOf_processStep_Flow
FUNCTION_BLOCK FB_ListOf_processStep_Flow  EXTENDS KOSTAL_TC3_Components_ListOf_Objects.FB_Base IMPLEMENTS I_ListOf_processStep_Flow, I_ListOf_processStep_Flow_CopyFrom, I_ListOf_processStep_Flow_Owner

VAR
	_Dummy	: FB_processStep_Flow;
END_VAR

//Overwrites the method in the base class with the real contents of the ListOf class.
METHOD PROTECTED  _deletePayLoad
VAR_INPUT
	pPayload	:	PVOID; 
END_VAR

VAR
	_p	: POINTER TO FB_processStep_Flow;
END_VAR

IF pPayload = 0  THEN	RETURN;	END_IF

_p:= pPayload;

__DELETE(_p);
END_METHOD

